// Device/Application/02_Devices/FB_RealCylinderGroup
FUNCTION_BLOCK FB_RealCylinderGroup
(* 模块说明：按料型选通的真实气缸组适配层（G2 侧挡用，300/450/600 三缸共用设备索引 10）。
   同一时刻只允许一个气缸下降，其余两个强制提升；回写与 FB_SimDevice 完全一致的接收/完成序号，
   使上层流程与互锁无需区分单缸、多缸或仿真。
   命令目标 lrTarget：0 = 三缸全部提升；300 / 450 / 600 = 对应料型气缸下降，其余两个提升。
   lrTarget 在 0..1 之间时按单缸旧语义映射：>0.5 视为「降到当前料型」，<=0.5 视为三缸全部提升。 *)
VAR_INPUT
	xUseReal : BOOL; (* TRUE 表示本编号由真实气缸组接管；FALSE 时三个阀全部失电且不响应任何命令。 *)
	xEnable : BOOL; (* 设备级使能，来自整机许可；FALSE 时阀失电并清序号。 *)
	xReset : BOOL; (* 故障复位上升沿；清锁存错误与序号。 *)
	xFaultHold : BOOL; (* 整机故障保持：TRUE 时三个阀立即失电，直到复位。 *)
	uiMaterialModel : UINT; (* 当前运行料型 300/450/600；旧语义 lrTarget>0.5 时降到本料型。 *)
	xSensorRetract1 : BOOL; (* 1 号缸（300）提升到位传感器原始电平，TRUE 表示该端有信号。 *)
	xSensorExtend1 : BOOL; (* 1 号缸（300）下降到位传感器原始电平。 *)
	xSensorRetract2 : BOOL; (* 2 号缸（450）提升到位传感器原始电平。 *)
	xSensorExtend2 : BOOL; (* 2 号缸（450）下降到位传感器原始电平。 *)
	xSensorRetract3 : BOOL; (* 3 号缸（600）提升到位传感器原始电平。 *)
	xSensorExtend3 : BOOL; (* 3 号缸（600）下降到位传感器原始电平。 *)
	xInvertSensors : BOOL; (* TRUE 表示六个传感器均为低电平有效，本层统一取反，不动上层。 *)
	xInvertValve : BOOL; (* TRUE 表示三个阀均为低电平使能；默认 FALSE，即高电平使能。 *)
	tSensorTimeout : TIME := T#3S; (* 六个传感器全部无信号达到该时间判为整组丢失，报 3004。 *)
	tTravelTimeout : TIME := T#10S; (* 命令发出后目标姿态未达成达到该时间判为动作超时，报 3005。 *)
	stConfig : ST_DeviceConfig; (* 行程范围，语义与仿真侧一致；组内气缸只使用 0/1 两端。 *)
	stCommand : ST_DeviceCommand; (* 上层统一设备命令，本层只响应 Position 的 0/300/450/600 目标。 *)
END_VAR
VAR_OUTPUT
	stStatus : ST_DeviceStatus; (* 与 FB_SimDevice 语义一致；目标缸下降到位 1.0，三缸全提 0.0，中间保持上次值。 *)
	aValve : ARRAY[1..3] OF BOOL; (* 三个阀的电气电平（已含 xInvertValve），直接接物理输出点；索引 1=300，2=450，3=600。 *)
	uiActiveBand : UINT; (* 当前实际下降的料型带号；0 表示三个缸都在提升位。 *)
END_VAR
VAR
	rtReset : R_TRIG; (* 复位上升沿。 *)
	tonNoSensor : TON; (* 六个传感器全部无信号的持续计时。 *)
	tonTravel : TON; (* 命令发出后等待到位的计时。 *)
	udiLastID : UDINT; (* 上次已接受的命令序号。 *)
	aRetract : ARRAY[1..3] OF BOOL; (* 取反处理后的三路提升信号。 *)
	aExtend : ARRAY[1..3] OF BOOL; (* 取反处理后的三路下降信号。 *)
	xAllRetract : BOOL; (* 三个缸都确认在提升位。 *)
	xPositionKnown : BOOL; (* 三缸姿态是否都已由传感器确立；未确立时 xReady 必须为 FALSE，防止上层把未知当成已提升。 *)
	xCmdValid : BOOL; (* 当前存在有效的保位命令，阀按此持续输出。 *)
	uiTargetBand : UINT; (* 有效命令期望下降的料型带号；0 表示三缸全部提升。 *)
	xTravelling : BOOL; (* 尚未确认到达命令要求的姿态。 *)
	i : INT; (* 本扫描数组遍历索引；含义及范围以当前 FOR 循环为准。 *)
END_VAR

rtReset(CLK := xReset);

(* ===== 1. 复位：只清错误与序号，姿态仍由传感器决定 ===== *)
IF xUseReal AND rtReset.Q THEN
	stStatus.xError := FALSE; stStatus.udiErrorID := 0;
	xCmdValid := FALSE; xTravelling := FALSE; udiLastID := 0; uiTargetBand := 0;
	stStatus.udiAcceptedID := 0; stStatus.udiCompletedID := 0;
	tonNoSensor(IN := FALSE);
	tonTravel(IN := FALSE);
END_IF

(* ===== 2. 传感器取反与逐缸姿态判定 ===== *)
aRetract[1] := xSensorRetract1 XOR xInvertSensors;
aExtend[1] := xSensorExtend1 XOR xInvertSensors;
aRetract[2] := xSensorRetract2 XOR xInvertSensors;
aExtend[2] := xSensorExtend2 XOR xInvertSensors;
aRetract[3] := xSensorRetract3 XOR xInvertSensors;
aExtend[3] := xSensorExtend3 XOR xInvertSensors;

(* 单缸两端同时有信号：传感器短路、磁环位置错或机械卡在中间，该缸姿态不可信，按 3003 暴露。
   逐缸判定而不是整组判定：只要有一个缸自相矛盾，整组位置就不可信。 *)
FOR i := 1 TO 3 DO
	IF aRetract[i] AND aExtend[i] THEN
		stStatus.xError := TRUE; stStatus.udiErrorID := 3003;
	END_IF
END_FOR

(* 三缸姿态是否都已确立：每个缸必须恰好一端有效，中间态或两端全无都算未确立。 *)
xAllRetract := aRetract[1] AND aRetract[2] AND aRetract[3];
xPositionKnown := TRUE;
FOR i := 1 TO 3 DO
	IF (NOT aRetract[i]) AND (NOT aExtend[i]) THEN xPositionKnown := FALSE; END_IF
END_FOR
IF stStatus.xError THEN xPositionKnown := FALSE; END_IF

(* 六个传感器全部无信号并持续 tSensorTimeout：判整组传感器丢失，报 3004。
   单缸丢失不在这里报，由 xPositionKnown 为 FALSE 阻断就绪，交给超时暴露，避免一缸调试刷整组报警。 *)
tonNoSensor(IN := xUseReal AND NOT aRetract[1] AND NOT aExtend[1]
	AND NOT aRetract[2] AND NOT aExtend[2]
	AND NOT aRetract[3] AND NOT aExtend[3], PT := tSensorTimeout);
IF tonNoSensor.Q AND NOT stStatus.xError THEN
	stStatus.xError := TRUE; stStatus.udiErrorID := 3004;
END_IF

(* ===== 3. 命令接收与保位判定 ===== *)
IF NOT xUseReal THEN
	(* 未接管：不驱动阀，也不发布就绪，避免被上层当成可用设备 *)
	xCmdValid := FALSE; xTravelling := FALSE; udiLastID := 0; uiTargetBand := 0;
	stStatus.xReady := FALSE; stStatus.xBusy := FALSE; stStatus.xActive := FALSE;
	stStatus.udiAcceptedID := 0; stStatus.udiCompletedID := 0;
ELSIF NOT xEnable OR stStatus.xError OR xFaultHold THEN
	(* 故障或整机故障保持时阀失电，不带错误继续动作 *)
	xCmdValid := FALSE; xTravelling := FALSE;
	stStatus.xReady := FALSE; stStatus.xBusy := FALSE; stStatus.xActive := FALSE;
ELSE
	stStatus.xReady := xEnable AND xPositionKnown;

	(* 新序号即新命令；姿态未确立时不接受，防止朝未知状态动作 *)
	IF (stCommand.udiID <> 0) AND (stCommand.udiID <> udiLastID)
		AND xEnable AND xPositionKnown AND NOT stStatus.xBusy THEN
		udiLastID := stCommand.udiID;
		stStatus.udiAcceptedID := udiLastID; stStatus.udiCompletedID := 0;
		CASE stCommand.eAction OF
		E_DeviceAction.Position:
			IF (stCommand.lrTarget > 0.5) AND (stCommand.lrTarget <= 1.0) THEN
				(* 单缸旧语义：1 = 降到当前料型；料型非法时报 2001，不猜一个缸去动作 *)
				IF (uiMaterialModel = 300) OR (uiMaterialModel = 450) OR (uiMaterialModel = 600) THEN
					uiTargetBand := uiMaterialModel;
				ELSE
					stStatus.xError := TRUE; stStatus.udiErrorID := 2001;
				END_IF
			ELSIF ABS(stCommand.lrTarget) < 0.01 THEN
				uiTargetBand := 0;
			ELSIF (ABS(stCommand.lrTarget - 300.0) < 0.01) THEN
				uiTargetBand := 300;
			ELSIF (ABS(stCommand.lrTarget - 450.0) < 0.01) THEN
				uiTargetBand := 450;
			ELSIF (ABS(stCommand.lrTarget - 600.0) < 0.01) THEN
				uiTargetBand := 600;
			ELSE
				(* 只支持 0 / 300 / 450 / 600，其它目标明确报错而不是静默不动 *)
				stStatus.xError := TRUE; stStatus.udiErrorID := 2001;
			END_IF
			IF NOT stStatus.xError THEN
				xCmdValid := TRUE;
				xTravelling := TRUE;
				stStatus.xBusy := TRUE;
			ELSE
				xCmdValid := FALSE;
			END_IF
		E_DeviceAction.Stop, E_DeviceAction.None:
			xCmdValid := FALSE; xTravelling := FALSE; uiTargetBand := 0;
			stStatus.udiAcceptedID := 0; stStatus.udiCompletedID := 0;
			udiLastID := 0;
		ELSE
			(* 气缸组没有连续运行、点动和回零，明确报错而不是静默不动 *)
			stStatus.xError := TRUE; stStatus.udiErrorID := 2001;
			xCmdValid := FALSE;
		END_CASE
	END_IF

	(* 命令被撤销或失能：立即取消保位，阀随之失电 *)
	IF (stCommand.eAction = E_DeviceAction.Stop) OR (stCommand.eAction = E_DeviceAction.None)
		OR NOT xEnable THEN
		xCmdValid := FALSE; xTravelling := FALSE;
		stStatus.xBusy := FALSE;
	END_IF

	(* 到位判定：目标缸下降到位，并且另外两个缸都在提升位，才算本次命令完成。
	   中间态（目标缸还没下去、或另一缸还没起来）都视为未完成，由超时兜底。 *)
	IF xCmdValid AND xPositionKnown THEN
		CASE uiTargetBand OF
		0:
			IF xAllRetract THEN
				IF xTravelling THEN stStatus.udiCompletedID := udiLastID; END_IF
				xTravelling := FALSE;
				stStatus.xBusy := FALSE;
			END_IF
		300:
			IF aExtend[1] AND aRetract[2] AND aRetract[3] THEN
				IF xTravelling THEN stStatus.udiCompletedID := udiLastID; END_IF
				xTravelling := FALSE;
				stStatus.xBusy := FALSE;
			END_IF
		450:
			IF aExtend[2] AND aRetract[1] AND aRetract[3] THEN
				IF xTravelling THEN stStatus.udiCompletedID := udiLastID; END_IF
				xTravelling := FALSE;
				stStatus.xBusy := FALSE;
			END_IF
		600:
			IF aExtend[3] AND aRetract[1] AND aRetract[2] THEN
				IF xTravelling THEN stStatus.udiCompletedID := udiLastID; END_IF
				xTravelling := FALSE;
				stStatus.xBusy := FALSE;
			END_IF
		END_CASE
	END_IF
END_IF

(* ===== 4. 位置反馈：只有确切在位才更新，中间态保持上次值 ===== *)
IF uiTargetBand = 0 THEN
	IF xAllRetract THEN stStatus.lrPosition := 0.0; END_IF
ELSIF uiTargetBand = 300 THEN
	IF aExtend[1] THEN stStatus.lrPosition := 1.0; END_IF
ELSIF uiTargetBand = 450 THEN
	IF aExtend[2] THEN stStatus.lrPosition := 1.0; END_IF
ELSIF uiTargetBand = 600 THEN
	IF aExtend[3] THEN stStatus.lrPosition := 1.0; END_IF
END_IF

(* 实际下降的料型：命令目标有效且该缸确实到位才报带号，避免阀已得电但没下去时谎报挡料就位 *)
uiActiveBand := 0;
IF (uiTargetBand = 300) AND aExtend[1] THEN uiActiveBand := 300; END_IF
IF (uiTargetBand = 450) AND aExtend[2] THEN uiActiveBand := 450; END_IF
IF (uiTargetBand = 600) AND aExtend[3] THEN uiActiveBand := 600; END_IF

(* ===== 5. 到位超时 ===== *)
tonTravel(IN := xUseReal AND xTravelling AND xCmdValid, PT := tTravelTimeout);
IF tonTravel.Q AND NOT stStatus.xError THEN
	stStatus.xError := TRUE; stStatus.udiErrorID := 3005;
	stStatus.xBusy := FALSE;
	xTravelling := FALSE;
END_IF

(* ===== 6. 阀输出：按保位命令持续输出，不是只在动作过程中输出；任何时刻最多一个缸下降 ===== *)
aValve[1] := FALSE; aValve[2] := FALSE; aValve[3] := FALSE;
IF xCmdValid AND xUseReal AND NOT stStatus.xError AND NOT xFaultHold THEN
	aValve[1] := (uiTargetBand = 300);
	aValve[2] := (uiTargetBand = 450);
	aValve[3] := (uiTargetBand = 600);
END_IF
IF xInvertValve THEN
	aValve[1] := NOT aValve[1]; aValve[2] := NOT aValve[2]; aValve[3] := NOT aValve[3];
END_IF

(* ===== 7. 收尾 ===== *)
stStatus.xReady := stStatus.xReady AND xUseReal AND NOT stStatus.xError;
stStatus.xActive := xCmdValid;
(* 气缸组没有回零动作，用「三缸姿态都已确立」代替，供整机统计已接管设备是否可信 *)
stStatus.xHomed := xUseReal AND xPositionKnown;

END_FUNCTION_BLOCK

// Device/Application/02_Devices/FB_RealSensor
FUNCTION_BLOCK FB_RealSensor
(* 模块说明：真实传感器（光电/接近开关）只读适配层。本块不驱动任何输出，只把原始电平
   去抖后发布成「到位」状态，使上层（自动送料判断、互锁、诊断）与仿真设备使用同一套接口。
   按料型/来料判断的是「有没有件」而不是「走到哪个位置」，所以姿态只有 0.0 / 1.0 两端：
   1.0 = 有料（光电被遮挡），0.0 = 无料。连续位置对传感器没有意义。 *)
VAR_INPUT
	xUseReal : BOOL; (* TRUE 表示本编号由真实传感器接管；FALSE 时不读物理点，也不发布就绪。 *)
	xEnable : BOOL; (* 设备级使能，来自整机许可；FALSE 时状态复位为无料且不发布就绪。 *)
	xReset : BOOL; (* 故障复位上升沿；清锁存错误。 *)
	xSensorRaw : BOOL; (* 传感器原始电平，TRUE 表示被遮挡（有料）。 *)
	xInvertSensor : BOOL; (* TRUE 表示接线为低电平有效（遮挡时读 FALSE），本层统一取反，不动上层。 *)
	tDebounce : TIME := T#20MS; (* 去抖时间：光电受粉尘、振动、反光影响会抖，短于该时间的跳变忽略。 *)
	tStuckTimeout : TIME := T#0MS; (* 常亮/常灭监视；0 表示不监视。料走完仍长时间有信号通常代表传感器卡死或反光。 *)
	stConfig : ST_DeviceConfig; (* 与其它设备一致的配置结构；传感器只用 lrInitialPosition 作初值，不使用行程字段。 *)
	stCommand : ST_DeviceCommand; (* 上层统一设备命令；传感器只响应被读请求，Position 目标被忽略。 *)
END_VAR
VAR_OUTPUT
	stStatus : ST_DeviceStatus; (* 与仿真侧语义一致；lrPosition 取 1.0 有料、0.0 无料。 *)
	xDetected : BOOL; (* 去抖后的最终信号，TRUE=有料。流程与互锁直接取用这个而不是原始点。 *)
	xRaw : BOOL; (* 取反处理后的原始电平（未去抖），供在线排查接线极性与抖动。 *)
END_VAR
VAR
	rtReset : R_TRIG; (* 复位上升沿。 *)
	tonDebounce : TON; (* 由 FALSE 变 TRUE 的去抖计时，到时才认「有料」。 *)
	tonClear : TON; (* 由 TRUE 变 FALSE 的去抖计时，到时才认「无料」。 *)
	tonStuck : TON; (* 长时间保持同一状态计时，用于常亮/常灭监视。 *)
	xStuckWindowClear : BOOL; (* 本扫描检测到电平跳变：清掉常亮/常灭计时窗口，重新开始计时。 *)
	xStable : BOOL; (* 去抖后的稳定值。 *)
	xLastRaw : BOOL; (* 上扫描取反后的原始电平，用于判断是否发生跳变并重置去抖计时。 *)
	xBooted : BOOL; (* 首次扫描标志，上电时直接用当前电平作初值，不等待去抖。 *)
END_VAR

rtReset(CLK := xReset);

(* ===== 1. 复位：只清错误，状态仍由传感器决定 ===== *)
IF xUseReal AND rtReset.Q THEN
	stStatus.xError := FALSE; stStatus.udiErrorID := 0;
	tonStuck(IN := FALSE);
END_IF

(* ===== 2. 极性处理：接线反了只改 xInvertSensor 一个参数，上层不受影响 ===== *)
xRaw := xSensorRaw XOR xInvertSensor;

(* ===== 3. 去抖：跳变后必须稳定 tDebounce 才改 xStable ===== *)
(* 用两个单稳计时而不是一个沿检测，是为了让"抖动期间保持上次稳定值"这件事显式可见：
   信号连续抖动时两个计时都不会到时，xStable 保持在最后一个稳定值上。 *)
xStuckWindowClear := (NOT xBooted) OR (xRaw <> xLastRaw);
IF xStuckWindowClear THEN
	tonDebounce(IN := FALSE);
	tonClear(IN := FALSE);
	IF NOT xBooted THEN
		(* 上电直接用当前电平作初值，避免开机 20ms 内把有料当无料 *)
		xStable := xRaw;
		xBooted := TRUE;
	END_IF
	xLastRaw := xRaw;
END_IF

IF xUseReal THEN
	IF xRaw THEN
		tonDebounce(IN := TRUE, PT := tDebounce);
		tonClear(IN := FALSE);
		IF tonDebounce.Q THEN xStable := TRUE; END_IF
	ELSE
		tonClear(IN := TRUE, PT := tDebounce);
		tonDebounce(IN := FALSE);
		IF tonClear.Q THEN xStable := FALSE; END_IF
	END_IF
END_IF

xDetected := xStable;

(* ===== 4. 常亮/常灭监视：料已走完却一直有信号，或本该有料却一直没有，都报出来 =====
   只监视"信号纹丝不动"这个可观测事实，不猜业务含义；阈值由 tStuckTimeout 给，0 表示关闭。 *)
tonStuck(IN := xUseReal AND (tStuckTimeout > T#0MS) AND NOT xStuckWindowClear, PT := tStuckTimeout);
IF tonStuck.Q AND NOT stStatus.xError THEN
	stStatus.xError := TRUE;
	(* 3006：持续有信号（常亮/反光/卡死）；3007：持续无信号（断线/被挡/未接通） *)
	IF xDetected THEN stStatus.udiErrorID := 3006;
	ELSE stStatus.udiErrorID := 3007; END_IF
END_IF

(* ===== 5. 状态发布：传感器没有动作请求，只要接管且使能就算就绪 ===== *)
stStatus.lrPosition := SEL(xDetected, 0.0, 1.0);
stStatus.xReady := xUseReal AND xEnable AND NOT stStatus.xError;
stStatus.xActive := xUseReal AND xDetected;
stStatus.xBusy := FALSE;
(* 传感器没有回零概念，用"已接管且状态可信"代替 *)
stStatus.xHomed := xUseReal AND xBooted;
stStatus.xRealActive := xUseReal;

END_FUNCTION_BLOCK

// Device/Application/04_Machine/FB_ManualControl
(* 模块说明：将手动按钮转为统一设备请求。点动松开即取消；定位与回零请求保持到本次完成；D6 不调度。 *)
FUNCTION_BLOCK FB_ManualControl
VAR_INPUT
	xEnable : BOOL; (* 手动模式且按钮释放联锁已满足时允许；未使能也同步按钮快照。 *)
	stReal : ST_RealDeviceSettings; (* 真实设备接管设置；真实编号的手动速度收紧到验证速度。 *)
	aManual : ARRAY[1..17] OF ST_ManualCommand; (* 各设备手动请求，索引 1..17；进入手动后先释放所有按钮再允许动作。 *)
END_VAR
VAR_IN_OUT
	aCommand : ARRAY[1..17] OF ST_DeviceCommand; (* 统一设备请求数组 1..17；子流程写请求，设备管理器执行。 *)
	aStatus : ARRAY[1..17] OF ST_DeviceStatus; (* 各设备的反馈数组 1..17，供判断忙、完成序号、故障和位置。 *)
	udiCounter : UDINT; (* 全机共享的动作序号计数器，通过引用传递；由 F_NextID 分配，0 不使用。 *)
END_VAR
VAR_OUTPUT
	uiRejectDevice : UINT; (* 本扫描最后一个手动拒绝设备索引；0 无，常见原因是冲突按钮或不支持该动作。 *)
END_VAR
VAR
	aPrev : ARRAY[1..17] OF ST_ManualCommand; (* 上扫描手动按钮快照；即使禁用仍更新，防止按住按钮切模式后被误作新上升沿。 *)
	aPending : ARRAY[1..17] OF ST_DeviceCommand; (* 手动定位或回零的锁存请求，直到本次命令完成；点动或运行优先时清除。 *)
	aRunID : ARRAY[1..17] OF UDINT; (* 各设备按住运行/点动时保持的序号，按钮释放后归零。 *)
	i : INT; (* 本扫描数组遍历索引；含义及范围以当前 FOR 循环为准。 *)
	lrVelocity : LREAL; (* 本扫描限幅后的手动速度，取绝对值限幅 0.1..100；反向点动时变为负值。 *)
	lrVelocityMax : LREAL; (* 本扫描速度上限；真实设备收紧到验证速度，防止全速冲出。 *)
	uiPressed : UINT; (* 本扫描该设备同时按下的手动按钮个数；大于 1 视为冲突并拒绝。 *)
END_VAR

(* 每扫描重新判断按钮冲突；无合法请求的设备由整机统一撤销动作。 *)
uiRejectDevice:=0;
FOR i:=1 TO 17 DO
    IF NOT xEnable THEN
        aPending[i].eAction:=E_DeviceAction.None;
        aRunID[i]:=0;
    ELSIF i<>6 THEN
        (* 先撤销本设备请求，只有命中合法按钮时才在下面重新写入。否则松开点动后，
           上一扫描的 Jog 会一直残留在共享请求数组里，真实轴靠 None/Stop 停止的逻辑永远等不到。 *)
        aCommand[i]:=F_Command(E_DeviceAction.None,0,0.0,0.0);
        (* 真实设备的手动速度上限由 lrManualVelocityMax 决定（默认 200）；实际速度取 aManual[i].lrVelocity 与之较小者。 *)
        lrVelocityMax:=100.0;
        IF stReal.axRealDevice[i] THEN
            (* 新字段在未重新初始化的旧下载里可能为 0；兜底 100，避免手动速度变 0 表现为不动作 *)
            lrVelocityMax:=100.0;
            IF stReal.lrManualVelocityMax>0.1 THEN lrVelocityMax:=LIMIT(0.1,stReal.lrManualVelocityMax,200.0); END_IF
        END_IF
        IF i=8 THEN
            (* D8 平台旋转轴（主轴）手动默认 3、限速 5；请求值超过上限时按默认 3 走，不要直接跳到 5。 *)
            lrVelocityMax:=5.0;
            lrVelocity:=3.0;
            IF ABS(aManual[i].lrVelocity)<=lrVelocityMax THEN
                lrVelocity:=LIMIT(0.1,ABS(aManual[i].lrVelocity),lrVelocityMax);
            END_IF
        ELSE
            lrVelocity:=LIMIT(0.1,ABS(aManual[i].lrVelocity),lrVelocityMax);
        END_IF
        (* 任意两个手动按钮同时按下都算冲突：正反点动、点动与定位/运行/回零、定位与运行/回零、运行与回零。 *)
        uiPressed:=0;
        IF aManual[i].xJogPositive THEN uiPressed:=uiPressed+1; END_IF
        IF aManual[i].xJogNegative THEN uiPressed:=uiPressed+1; END_IF
        IF aManual[i].xMove THEN uiPressed:=uiPressed+1; END_IF
        IF aManual[i].xRun THEN uiPressed:=uiPressed+1; END_IF
        IF aManual[i].xHome THEN uiPressed:=uiPressed+1; END_IF
        IF uiPressed>1 THEN
            uiRejectDevice:=INT_TO_UINT(i); aPending[i].eAction:=E_DeviceAction.None;
        (* 点动电平控制，只支持 D2/D4/D5/D7/D8；速度符号决定方向，松开后不保持点动。 *)
        ELSIF aManual[i].xJogPositive OR aManual[i].xJogNegative THEN
            aPending[i].eAction:=E_DeviceAction.None;
            IF aRunID[i]=0 THEN aRunID[i]:=F_NextID(udiCounter); END_IF
            IF aManual[i].xJogNegative THEN lrVelocity:=-lrVelocity; END_IF
            IF (i=2) OR (i=4) OR (i=5) OR (i=7) OR (i=8) THEN
                aCommand[i]:=F_Command(E_DeviceAction.Jog,aRunID[i],0.0,lrVelocity);
            ELSE uiRejectDevice:=INT_TO_UINT(i);
            END_IF
        (* 连续运行电平控制，仅允许皮带、盘刀、喷油和吹气；盘刀接真实轴后走 FB_RealAxis 的 Run 相位。 *)
        ELSIF aManual[i].xRun THEN
            aPending[i].eAction:=E_DeviceAction.None;
            IF (i=1) OR (i=3) OR (i=13) OR (i=14) THEN
                IF aRunID[i]=0 THEN aRunID[i]:=F_NextID(udiCounter); END_IF
                aCommand[i]:=F_Command(E_DeviceAction.Run,aRunID[i],0.0,lrVelocity);
            ELSE uiRejectDevice:=INT_TO_UINT(i);
            END_IF
        (* 回零：上升沿锁存一次请求，之后每扫描重发直到完成；真实轴 D2/D8，D4 为仿真但保留入口。
           D3 盘刀是连续旋转主轴，只做 Run 不做回零，因此不在本白名单内。
           这里不能像点动那样在分支开头清 aPending —— 回零是保持型动作，清了就只剩一个扫描周期，
           设备刚接收就会被下一扫描的 None 撤销，表现为「下发了但不动」。 *)
        ELSIF aManual[i].xHome THEN
            aRunID[i]:=0;
            IF (i=2) OR (i=4) OR (i=8) THEN
                IF NOT aPrev[i].xHome THEN
                    aPending[i]:=F_Command(E_DeviceAction.Home,F_NextID(udiCounter),0.0,0.0);
                END_IF
                IF aPending[i].eAction<>E_DeviceAction.None THEN
                    aCommand[i]:=aPending[i];
                    IF F_Done(aStatus[i],aPending[i].udiID) THEN aPending[i].eAction:=E_DeviceAction.None; END_IF
                END_IF
            ELSE
                (* 不支持的编号：清掉可能从定位继承来的请求，避免继续执行上一个动作。 *)
                uiRejectDevice:=INT_TO_UINT(i);
                aPending[i].eAction:=E_DeviceAction.None;
            END_IF
        ELSE
            aRunID[i]:=0;
            (* 定位仅在按钮上升沿锁存目标和序号，然后持续等待本次完成。 *)
            IF aManual[i].xMove AND NOT aPrev[i].xMove THEN
                IF (i<>1) AND (i<>3) AND (i<>13) AND (i<>14) THEN
                    aPending[i]:=F_Command(E_DeviceAction.Position,F_NextID(udiCounter),aManual[i].lrTarget,lrVelocity);
                ELSE uiRejectDevice:=INT_TO_UINT(i);
                END_IF
            END_IF
            IF aPending[i].eAction<>E_DeviceAction.None THEN
                aCommand[i]:=aPending[i];
                IF F_Done(aStatus[i],aPending[i].udiID) THEN aPending[i].eAction:=E_DeviceAction.None; END_IF
            END_IF
        END_IF
    END_IF
    (* 禁用时仍同步按钮快照，避免按住定位按钮切入手动后产生虚假的新上升沿。 *)
    aPrev[i]:=aManual[i];
END_FOR

END_FUNCTION_BLOCK

// Device/Application/02_Devices/F_Command
(* 模块说明：组装设备命令，不执行运动。由设备管理器和对应设备功能块实际处理。 *)
FUNCTION F_Command : ST_DeviceCommand
VAR_INPUT
    eAction : E_DeviceAction; (* 动作类型：无请求、定位、连续运行、点动或停止，见 E_DeviceAction。 *)
    udiID : UDINT; (* 本次命令序号，0 无效；发起新定位时换新序号。 *)
    lrTarget : LREAL; (* 目标工程位置；气缸使用约定的 0/1 端点，连续运行和点动不使用该位置。 *)
    lrVelocity : LREAL; (* 请求速度，单位随设备工程单位定义；尚未完成实机标定。 *)
END_VAR

(* 只复制字段形成结构体，不等待动作、不直接访问物理设备。 *)
F_Command.eAction := eAction;
F_Command.udiID := udiID;
F_Command.lrTarget := lrTarget;
F_Command.lrVelocity := lrVelocity;

END_FUNCTION

// Device/Application/02_Devices/F_NextID
(* 模块说明：生成本次动作的非零序号。计数到最大值后回到 1，用于排除上一步残留的完成反馈。 *)
FUNCTION F_NextID : UDINT
VAR_IN_OUT
    udiCounter : UDINT; (* 全机共享的动作序号计数器，通过引用传递；由 F_NextID 分配，0 不使用。 *)
END_VAR

(* 最大值之后回到 1，跳过无效序号 0；同一机台所有流程共享该计数器。 *)
IF udiCounter = 16#FFFFFFFF THEN udiCounter := 1;
ELSE udiCounter := udiCounter + 1;
END_IF
F_NextID := udiCounter;

END_FUNCTION

// Device/Application/02_Devices/F_Done
(* 模块说明：只有设备完成序号等于本次命令序号、无忙且无故障，才返回动作完成。 *)
FUNCTION F_Done : BOOL
VAR_INPUT
    stStatus : ST_DeviceStatus; (* 本模块对外发布的状态；字段含义见其数据类型。 *)
    udiID : UDINT; (* 本次命令序号，0 无效；发起新定位时换新序号。 *)
END_VAR

(* 完成必须匹配本次请求；历史 Done 或仅 Busy=FALSE 都不足以作为本步完成条件。 *)
F_Done := (udiID <> 0) AND (stStatus.udiCompletedID = udiID)
    AND NOT stStatus.xBusy AND NOT stStatus.xError;

END_FUNCTION

// Device/Application/04_Machine/FB_AutoCycle
(* 模块说明：自动主状态机。只组织工序并提出请求，设备执行由整机统一调用；送料等料允许长期等待。 *)
FUNCTION_BLOCK FB_AutoCycle
VAR_INPUT
    xRun : BOOL; (* 自动工序运行许可，整机 Automatic 时保持 TRUE；撤销立即复位主流程。 *)
    xContinuous : BOOL; (* TRUE 连续循环；FALSE 在当前完整循环结束后回到就绪。 *)
    xMaterialAtLength : BOOL; (* 定长光电到位状态；自动送料须先离开再到位，并满足 D5 下降。 *)
    stRecipe : ST_Recipe; (* 待校验配方或上层传入的运行配方，字段含义见 ST_Recipe。 *)
END_VAR
VAR_IN_OUT
    aCommand : ARRAY[1..17] OF ST_DeviceCommand; (* 统一设备请求数组 1..17；子流程写请求，设备管理器执行。 *)
    aStatus : ARRAY[1..17] OF ST_DeviceStatus; (* 各设备的反馈数组 1..17，供判断忙、完成序号、故障和位置。 *)
    udiCounter : UDINT; (* 全机共享的动作序号计数器，通过引用传递；由 F_NextID 分配，0 不使用。 *)
END_VAR
VAR_OUTPUT
    eStep : E_AutoStep; (* 自动主工序当前状态，见 E_AutoStep。 *)
    xDone : BOOL; (* 整循环完成的单扫描脉冲；机械手等三路收尾全部结束后才产生。 *)
    xError : BOOL; (* 本设备或本子流程发生故障；具体原因见对应错误码。 *)
    udiErrorID : UDINT; (* 非法主步骤为 4800；主步超时为 4800+步号；步骤守护失败为 4800+步号+1，见下方守护表；支线错误则向上传递。 *)
    uiClearLengthStep : UINT; (* 避让支线 P 的当前步骤：10 升起 D5，20 移开 D4，1000 完成。 *)
    uiClearTransferStep : UINT; (* 避让支线 Q 当前步骤：10 降 G4，20 松 G3，30 降 G2，1000 完成。 *)
    uiPostStep : UINT; (* 收尾总步骤：10 抬刀，20 抬压，30 等待三路完成，1000 结束。 *)
    uiReturnKnifeStep : UINT; (* 收尾支线 A：10 喷油，20 D2 回刀，1000 完成。 *)
    uiUnloadStep : UINT; (* 机械手移料支线 B 步骤，10..110 每步加 10，1000 完成；详见 FB_Unload。 *)
    uiResetLengthStep : UINT; (* 收尾支线 C：10 D4 定位，20 D5 下降，30 确认下降，1000 完成。 *)
END_VAR
VAR
    ePrevStep : E_AutoStep := E_AutoStep.Fault; (* 上扫描主工序状态，用于产生步骤入口标志。 *)
    udiToken : UDINT; (* 本步骤专用动作序号；同一步中的设备共用该号，以排除旧完成信号。 *)
    udiSpindleToken : UDINT; (* 盘刀运行命令序号，切割过程中保持该号，避免重复重启盘刀命令。 *)
    udiPressToken : UDINT; (* G1 下压保位序号；PressDown 入口分配，后续步骤持续用该号重发，保证单电控阀不断电。 *)
    udiKnifeToken : UDINT; (* G9 下刀保位序号；KnifeDown 入口分配，同上。 *)
    xEntry : BOOL; (* 本扫描为新步骤入口；用于分配新序号并复位步骤超时计时。 *)
    xSawSensorClear : BOOL; (* 本轮送料已观察到光电离开；须先有该标志再接受新到位，防止残留信号触发。 *)
    tonStep : TON; (* 步骤超时定时器；进入新步骤时复位，超时错误码由模块及当前步号组成。 *)
    tStepLimit : TIME; (* 本扫描用的步骤超时值：切割步取 tCutTimeout，其余取 tStepTimeout。 *)
    xGuardOK : BOOL; (* 步骤守护判据：当前步依赖的前提是否仍满足，FALSE 时立即报错退出，不等步超时。 *)
    fbClear : FB_ClearanceUnit; (* 切割前两路并行避让流程。 *)
    fbPost : FB_PostCut; (* 切割后抬刀、抬压及三路收尾流程。 *)
END_VAR

(* 完成标志每扫描先清零；本流程在许可撤销后复位，不保留中断点续跑。 *)
xDone := FALSE;
IF NOT xRun THEN eStep:=E_AutoStep.Idle; xError:=FALSE; udiErrorID:=0; xSawSensorClear:=FALSE; END_IF
(* 进入新步骤才换新动作序号，同一步持续保持请求，防止反复启动。 *)
xEntry := eStep <> ePrevStep;
IF xEntry THEN udiToken := F_NextID(udiCounter); END_IF
ePrevStep := eStep;
(* 送料等料不计步骤超时；其余执行步按运行配方监控。
   切割步单独用 tCutTimeout：走刀行程长，和其它单动作步共用一个 30 秒很容易误超时。 *)
tStepLimit := stRecipe.tStepTimeout;
IF eStep = E_AutoStep.Cutting THEN tStepLimit := stRecipe.tCutTimeout; END_IF
tonStep(IN:=xRun AND NOT xEntry AND (eStep<>E_AutoStep.Idle)
    AND (eStep<>E_AutoStep.FeedWait) AND (eStep<>E_AutoStep.Complete)
    AND (eStep<>E_AutoStep.Fault),PT:=tStepLimit);
IF xRun AND NOT xError THEN
CASE eStep OF
(* 待机转入送料；没有直接跳到切割。 *)
E_AutoStep.Idle: eStep:=E_AutoStep.FeedWait;
(* D1 送料并正常等料；光电须先离开再到位，且 D5 必须在下降端。 *)
E_AutoStep.FeedWait:
    IF xEntry THEN xSawSensorClear:=FALSE; END_IF
    IF NOT xMaterialAtLength THEN xSawSensorClear:=TRUE; END_IF
    aCommand[1]:=F_Command(E_DeviceAction.Run,udiToken,0.0,stRecipe.lrBeltVelocity);
    IF xSawSensorClear AND xMaterialAtLength AND F_At(aStatus[5],1.0) THEN eStep:=E_AutoStep.StopFeed; END_IF
(* 本步不再给 D1 运行请求，整机周期清空请求后等待皮带非运行、非忙。 *)
E_AutoStep.StopFeed:
    IF NOT aStatus[1].xActive AND NOT aStatus[1].xBusy THEN eStep:=E_AutoStep.Push; END_IF
(* G3 侧推到位；只认本次 udiToken 对应的完成。 *)
E_AutoStep.Push:
    aCommand[11]:=F_Command(E_DeviceAction.Position,udiToken,1.0,stRecipe.lrPositionVelocity);
    IF F_Done(aStatus[11],udiToken) THEN eStep:=E_AutoStep.Clearance; END_IF
(* 并行调用定长避让 P 和输送机构避让 Q，两路都完成后旋转平台。 *)
E_AutoStep.Clearance:
    IF fbClear.xDone THEN eStep:=E_AutoStep.Rotate; END_IF
(* D8 旋转到 lrRotateAngle，必须在 G1 下压之前完成。 *)
E_AutoStep.Rotate:
    aCommand[8]:=F_Command(E_DeviceAction.Position,udiToken,stRecipe.lrRotateAngle,stRecipe.lrPositionVelocity);
    IF F_Done(aStatus[8],udiToken) THEN eStep:=E_AutoStep.PressDown; END_IF
(* G1 下压到位。 *)
E_AutoStep.PressDown:
    IF xEntry THEN udiPressToken:=udiToken; END_IF
    aCommand[9]:=F_Command(E_DeviceAction.Position,udiPressToken,1.0,stRecipe.lrPositionVelocity);
    IF F_Done(aStatus[9],udiPressToken) THEN eStep:=E_AutoStep.SpindleOn; END_IF
(* D3 盘刀先转起来，转稳了再下刀；此时刀还没下来，G1 保持压紧。 *)
E_AutoStep.SpindleOn:
    udiSpindleToken:=udiToken;
    aCommand[9]:=F_Command(E_DeviceAction.Position,udiPressToken,1.0,stRecipe.lrPositionVelocity);
    aCommand[3]:=F_Command(E_DeviceAction.Run,udiSpindleToken,0.0,stRecipe.lrSpindleVelocity);
    IF F_Done(aStatus[3],udiSpindleToken) AND aStatus[3].xActive THEN eStep:=E_AutoStep.KnifeDown; END_IF
(* G9 盘刀下降到位；下降全程 D3 保持运行。 *)
E_AutoStep.KnifeDown:
    IF xEntry THEN udiKnifeToken:=udiToken; END_IF
    aCommand[9]:=F_Command(E_DeviceAction.Position,udiPressToken,1.0,stRecipe.lrPositionVelocity);
    aCommand[3]:=F_Command(E_DeviceAction.Run,udiSpindleToken,0.0,stRecipe.lrSpindleVelocity);
    aCommand[17]:=F_Command(E_DeviceAction.Position,udiKnifeToken,1.0,stRecipe.lrPositionVelocity);
    IF F_Done(aStatus[17],udiKnifeToken) THEN eStep:=E_AutoStep.Cutting; END_IF
(* 保持 D3 运行，G6 吹气，D2 走到回刀起点加切割长度；以 D2 到位作为切割完成。 *)
E_AutoStep.Cutting:
    aCommand[9]:=F_Command(E_DeviceAction.Position,udiPressToken,1.0,stRecipe.lrPositionVelocity);
    aCommand[17]:=F_Command(E_DeviceAction.Position,udiKnifeToken,1.0,stRecipe.lrPositionVelocity);
    aCommand[3]:=F_Command(E_DeviceAction.Run,udiSpindleToken,0.0,stRecipe.lrSpindleVelocity);
    aCommand[14]:=F_Command(E_DeviceAction.Run,udiToken,0.0,0.0);
    aCommand[2]:=F_Command(E_DeviceAction.Position,udiToken,stRecipe.lrCutHome+stRecipe.lrCutLength,stRecipe.lrCutVelocity);
    IF F_Done(aStatus[2],udiToken) THEN eStep:=E_AutoStep.StopCut; END_IF
(* 撤销 D3/G6 运行请求，等待盘刀停止且吹气关闭后收尾。 *)
E_AutoStep.StopCut:
    aCommand[9]:=F_Command(E_DeviceAction.Position,udiPressToken,1.0,stRecipe.lrPositionVelocity);
    aCommand[17]:=F_Command(E_DeviceAction.Position,udiKnifeToken,1.0,stRecipe.lrPositionVelocity);
    IF NOT aStatus[3].xActive AND NOT aStatus[3].xBusy AND NOT aStatus[14].xActive THEN eStep:=E_AutoStep.PostCut; END_IF
(* 先抬刀再抬压，随后三支线同步执行；全部结束才完成本轮。 *)
E_AutoStep.PostCut:
    IF fbPost.xDone THEN eStep:=E_AutoStep.Complete; END_IF
(* 只在进入本步时输出一次完成脉冲；连续模式返回送料，单循环由整机回到 Ready。 *)
E_AutoStep.Complete:
    xDone:=xEntry;
    IF xContinuous THEN eStep:=E_AutoStep.FeedWait; END_IF
(* 保留流程错误状态；整机退出自动后才复位此流程。 *)
E_AutoStep.Fault: xError:=TRUE;
ELSE xError:=TRUE; udiErrorID:=4800;
END_CASE
(* ===== 步骤守护表 =====
   只判前提，不判目标：目标是本步自己要去达成的东西，由各步的 F_Done 判完成；
   这里判的是这一步所依赖的前提还在不在。前提在进入该步时就已成立，
   之后必须一直保持，一旦丢失立即报错退出，不再干等 tonStep 超时才发现。
   每个步骤都要在下面有明确交代，无守护也要写出来，避免以后分不清
   是真的不需要还是漏掉了。新增步骤时先到这里补一行。
   错误码约定：4800 + 步号 + 1，例 SpindleOn=4881、Cutting=4891。
   这里不主动发 Stop：报错后本流程转 Fault，下一扫描不再提出任何请求，
   设备管理器收到 None 即停止，轴走 MC_Stop，气缸阀失电。 *)
xGuardOK := TRUE;
CASE eStep OF
(* 无守护：要么在等外部条件，要么本步本身就在建立条件。 *)
E_AutoStep.Idle, E_AutoStep.FeedWait, E_AutoStep.StopFeed,
E_AutoStep.Push, E_AutoStep.Clearance, E_AutoStep.Rotate,
E_AutoStep.PressDown, E_AutoStep.StopCut,
E_AutoStep.PostCut, E_AutoStep.Complete, E_AutoStep.Fault:
    xGuardOK := TRUE;

(* 起盘刀前：只要已压紧；此时刀还没下来，不判下刀。 *)
E_AutoStep.SpindleOn:
    xGuardOK := F_At(aStatus[9],1.0);

(* 下刀期间：压紧且盘刀必须已经在转，不能拿一把没转的刀往下扎。 *)
E_AutoStep.KnifeDown:
    xGuardOK := F_At(aStatus[9],1.0) AND aStatus[3].xActive;

(* 切割全程：压紧、下刀、盘刀运行三者都必须保持。 *)
E_AutoStep.Cutting:
    xGuardOK := F_At(aStatus[9],1.0) AND F_At(aStatus[17],1.0) AND aStatus[3].xActive;
END_CASE
IF NOT xGuardOK THEN
    xError := TRUE;
    udiErrorID := 4800 + TO_UDINT(eStep) + 1;
END_IF
IF tonStep.Q THEN xError:=TRUE; udiErrorID:=4800+TO_UDINT(eStep); END_IF
END_IF
(* 子功能块必须每扫描调用，包括失能时复位；上方状态判断看到的是此前反馈。 *)
fbClear(xExecute:=xRun AND (eStep=E_AutoStep.Clearance),stRecipe:=stRecipe,aCommand:=aCommand,aStatus:=aStatus,udiCounter:=udiCounter);
fbPost(xExecute:=xRun AND (eStep=E_AutoStep.PostCut),stRecipe:=stRecipe,aCommand:=aCommand,aStatus:=aStatus,udiCounter:=udiCounter);
(* 任一支线错误向主流程上报；所有设备请求还须经过整机统一互锁。 *)
IF fbClear.xError OR fbPost.xError THEN xError:=TRUE; udiErrorID:=MAX(fbClear.udiErrorID,fbPost.udiErrorID); END_IF
IF xError THEN eStep:=E_AutoStep.Fault; END_IF
uiClearLengthStep:=fbClear.uiLengthStep; uiClearTransferStep:=fbClear.uiTransferStep;
uiPostStep:=fbPost.uiStep; uiReturnKnifeStep:=fbPost.uiKnifeStep;
uiUnloadStep:=fbPost.uiUnloadStep; uiResetLengthStep:=fbPost.uiLengthStep;

END_FUNCTION_BLOCK

// Device/Application/03_Units/FB_Unload
(* 模块说明：收尾支线 B：机械手移料。后退、下降、最终回位是三个独立动作，全部完成后才允许下一轮送料。 *)
FUNCTION_BLOCK FB_Unload
VAR_INPUT
    xExecute : BOOL; (* 子流程执行许可；须保持到完成，清 FALSE 复位该流程步骤和错误。 *)
    stRecipe : ST_Recipe; (* 待校验配方或上层传入的运行配方，字段含义见 ST_Recipe。 *)
END_VAR
VAR_IN_OUT
    aCommand : ARRAY[1..17] OF ST_DeviceCommand; (* 统一设备请求数组 1..17；子流程写请求，设备管理器执行。 *)
    aStatus : ARRAY[1..17] OF ST_DeviceStatus; (* 各设备的反馈数组 1..17，供判断忙、完成序号、故障和位置。 *)
    udiCounter : UDINT; (* 全机共享的动作序号计数器，通过引用传递；由 F_NextID 分配，0 不使用。 *)
END_VAR
VAR_OUTPUT
    xDone : BOOL; (* 本子流程完成标志；执行许可撤销后复位。 *)
    xError : BOOL; (* 本设备或本子流程发生故障；具体原因见对应错误码。 *)
    udiErrorID : UDINT; (* 非法步骤码 4400；动作超时码=4400+uiStep，可据此定位本支线等待点。 *)
    uiStep : UINT; (* 当前子步骤：0 待机，10/20/... 执行动作，1000 完成；切勿在线强制跳步。 *)
END_VAR
VAR
    uiPrevStep : UINT := 65535; (* 上扫描步骤，用于判断本扫描是否刚进入新步骤。 *)
    udiToken : UDINT; (* 本步骤专用动作序号；同一步中的设备共用该号，以排除旧完成信号。 *)
    xEntry : BOOL; (* 本扫描为新步骤入口；用于分配新序号并复位步骤超时计时。 *)
    tonStep : TON; (* 步骤超时定时器；进入新步骤时复位，超时错误码由模块及当前步号组成。 *)
    tonSpray : TON; (* 通用子流程模板的喷油定时器，只有 FB_ReturnKnife 用其完成条件。 *)
END_VAR

(* 执行许可撤销即复位；步骤入口换新序号，每步等待本次动作完成，超时码=模块基码+步号。 *)
IF NOT xExecute THEN uiStep := 0; xError := FALSE; udiErrorID := 0; END_IF;
xEntry := uiStep <> uiPrevStep;
IF xEntry THEN udiToken := F_NextID(udiCounter); END_IF;
uiPrevStep := uiStep;
tonStep(IN := xExecute AND (uiStep > 0) AND (uiStep < 1000) AND NOT xEntry, PT := stRecipe.tStepTimeout);
tonSpray(IN := xExecute AND (uiStep = 10) AND aStatus[13].xActive, PT := stRecipe.tSpray);
IF xExecute AND NOT xError THEN
CASE uiStep OF
0: (* 待机；许可有效时进入首个动作。 *) uiStep := 10;
10: (* B010 侧挡 G2 提升。 *)
aCommand[10] := F_Command(E_DeviceAction.Position, udiToken, 0.0, stRecipe.lrPositionVelocity);
IF F_Done(aStatus[10], udiToken) THEN uiStep := 20; END_IF;
20: (* B020 流利条 G4 提升。 *)
aCommand[12] := F_Command(E_DeviceAction.Position, udiToken, 1.0, stRecipe.lrPositionVelocity);
IF F_Done(aStatus[12], udiToken) THEN uiStep := 30; END_IF;
30: (* B030 机械手 G7 提升。 *)
aCommand[15] := F_Command(E_DeviceAction.Position, udiToken, 1.0, stRecipe.lrPositionVelocity);
IF F_Done(aStatus[15], udiToken) THEN uiStep := 40; END_IF;
40: (* B040 夹爪 G8 打开，准备前进取料。 *)
aCommand[16] := F_Command(E_DeviceAction.Position, udiToken, 0.0, stRecipe.lrPositionVelocity);
IF F_Done(aStatus[16], udiToken) THEN uiStep := 50; END_IF;
50: (* B050 机械手 D7 前进到取料位置 lrGripperFront。 *)
aCommand[7] := F_Command(E_DeviceAction.Position, udiToken, stRecipe.lrGripperFront, stRecipe.lrPositionVelocity);
IF F_Done(aStatus[7], udiToken) THEN uiStep := 60; END_IF;
60: (* B060 夹爪 G8 夹紧，确认后才拉料。 *)
aCommand[16] := F_Command(E_DeviceAction.Position, udiToken, 1.0, stRecipe.lrPositionVelocity);
IF F_Done(aStatus[16], udiToken) THEN uiStep := 70; END_IF;
70: (* B070 机械手 D7 拉料到 lrGripperPull。 *)
aCommand[7] := F_Command(E_DeviceAction.Position, udiToken, stRecipe.lrGripperPull, stRecipe.lrPositionVelocity);
IF F_Done(aStatus[7], udiToken) THEN uiStep := 80; END_IF;
80: (* B080 夹爪 G8 打开，释放移走的料。 *)
aCommand[16] := F_Command(E_DeviceAction.Position, udiToken, 0.0, stRecipe.lrPositionVelocity);
IF F_Done(aStatus[16], udiToken) THEN uiStep := 90; END_IF;
90: (* B090 保持机械手抬升，D7 后退至 lrGripperBack；此时不是最终回位。 *)
aCommand[7] := F_Command(E_DeviceAction.Position, udiToken, stRecipe.lrGripperBack, stRecipe.lrPositionVelocity);
IF F_Done(aStatus[7], udiToken) THEN uiStep := 100; END_IF;
100: (* B100 后退到位后，G7 下降。 *)
aCommand[15] := F_Command(E_DeviceAction.Position, udiToken, 0.0, stRecipe.lrPositionVelocity);
IF F_Done(aStatus[15], udiToken) THEN uiStep := 110; END_IF;
110: (* B110 下降到位后，D7 再回 lrGripperHome；本支线结束前不允许送料。 *)
aCommand[7] := F_Command(E_DeviceAction.Position, udiToken, stRecipe.lrGripperHome, stRecipe.lrPositionVelocity);
IF F_Done(aStatus[7], udiToken) THEN uiStep := 1000; END_IF;
1000: (* 本支线完成，保持至 xExecute 撤销。 *) ;
ELSE xError := TRUE; udiErrorID := 4400;
END_CASE;
IF tonStep.Q THEN xError := TRUE; udiErrorID := 4400 + UINT_TO_UDINT(uiStep); END_IF;
END_IF;
xDone := xExecute AND (uiStep = 1000) AND NOT xError;

END_FUNCTION_BLOCK

// Device/Application/03_Units/FB_ReturnKnife
(* 模块说明：收尾支线 A：G5 喷油到设定时间，再令 D2 回刀。喷油仅在第一步保持请求。 *)
FUNCTION_BLOCK FB_ReturnKnife
VAR_INPUT
    xExecute : BOOL; (* 子流程执行许可；须保持到完成，清 FALSE 复位该流程步骤和错误。 *)
    stRecipe : ST_Recipe; (* 待校验配方或上层传入的运行配方，字段含义见 ST_Recipe。 *)
END_VAR
VAR_IN_OUT
    aCommand : ARRAY[1..17] OF ST_DeviceCommand; (* 统一设备请求数组 1..17；子流程写请求，设备管理器执行。 *)
    aStatus : ARRAY[1..17] OF ST_DeviceStatus; (* 各设备的反馈数组 1..17，供判断忙、完成序号、故障和位置。 *)
    udiCounter : UDINT; (* 全机共享的动作序号计数器，通过引用传递；由 F_NextID 分配，0 不使用。 *)
END_VAR
VAR_OUTPUT
    xDone : BOOL; (* 本子流程完成标志；执行许可撤销后复位。 *)
    xError : BOOL; (* 本设备或本子流程发生故障；具体原因见对应错误码。 *)
    udiErrorID : UDINT; (* 非法步骤码 4300；动作超时码=4300+uiStep，可据此定位本支线等待点。 *)
    uiStep : UINT; (* 当前子步骤：0 待机，10/20/... 执行动作，1000 完成；切勿在线强制跳步。 *)
END_VAR
VAR
    uiPrevStep : UINT := 65535; (* 上扫描步骤，用于判断本扫描是否刚进入新步骤。 *)
    udiToken : UDINT; (* 本步骤专用动作序号；同一步中的设备共用该号，以排除旧完成信号。 *)
    xEntry : BOOL; (* 本扫描为新步骤入口；用于分配新序号并复位步骤超时计时。 *)
    tonStep : TON; (* 步骤超时定时器；进入新步骤时复位，超时错误码由模块及当前步号组成。 *)
    tonSpray : TON; (* 通用子流程模板的喷油定时器，只有 FB_ReturnKnife 用其完成条件。 *)
END_VAR

(* 执行许可撤销即复位；步骤入口换新序号，每步等待本次动作完成，超时码=模块基码+步号。 *)
IF NOT xExecute THEN uiStep := 0; xError := FALSE; udiErrorID := 0; END_IF;
xEntry := uiStep <> uiPrevStep;
IF xEntry THEN udiToken := F_NextID(udiCounter); END_IF;
uiPrevStep := uiStep;
tonStep(IN := xExecute AND (uiStep > 0) AND (uiStep < 1000) AND NOT xEntry, PT := stRecipe.tStepTimeout);
tonSpray(IN := xExecute AND (uiStep = 10) AND aStatus[13].xActive, PT := stRecipe.tSpray);
IF xExecute AND NOT xError THEN
CASE uiStep OF
0: (* 待机；许可有效时进入首个动作。 *) uiStep := 10;
10: (* A010 G5 喷油并等待 tSpray；喷油建立后才开始计时。 *)
aCommand[13] := F_Command(E_DeviceAction.Run, udiToken, 0.0, 0.0);
IF tonSpray.Q THEN uiStep := 20; END_IF;
20: (* A020 结束喷油请求，D2 回到 lrCutHome，等待到位。 *)
aCommand[2] := F_Command(E_DeviceAction.Position, udiToken, stRecipe.lrCutHome, stRecipe.lrReturnVelocity);
IF F_Done(aStatus[2], udiToken) THEN uiStep := 1000; END_IF;
1000: (* 本支线完成，保持至 xExecute 撤销。 *) ;
ELSE xError := TRUE; udiErrorID := 4300;
END_CASE;
IF tonStep.Q THEN xError := TRUE; udiErrorID := 4300 + UINT_TO_UDINT(uiStep); END_IF;
END_IF;
xDone := xExecute AND (uiStep = 1000) AND NOT xError;

END_FUNCTION_BLOCK

// Device/Application/03_Units/FB_ClearanceUnit
(* 模块说明：并行执行 P/Q 两路避让；两路都完成才继续，任一路故障向主流程报告。 *)
FUNCTION_BLOCK FB_ClearanceUnit
VAR_INPUT
    xExecute : BOOL; (* 子流程执行许可；须保持到完成，清 FALSE 复位该流程步骤和错误。 *)
    stRecipe : ST_Recipe; (* 待校验配方或上层传入的运行配方，字段含义见 ST_Recipe。 *)
END_VAR
VAR_IN_OUT
    aCommand : ARRAY[1..17] OF ST_DeviceCommand; (* 统一设备请求数组 1..17；子流程写请求，设备管理器执行。 *)
    aStatus : ARRAY[1..17] OF ST_DeviceStatus; (* 各设备的反馈数组 1..17，供判断忙、完成序号、故障和位置。 *)
    udiCounter : UDINT; (* 全机共享的动作序号计数器，通过引用传递；由 F_NextID 分配，0 不使用。 *)
END_VAR
VAR_OUTPUT
    xDone : BOOL; (* 本子流程完成标志；执行许可撤销后复位。 *)
    xError : BOOL; (* 本设备或本子流程发生故障；具体原因见对应错误码。 *)
    udiErrorID : UDINT; (* 错误码；0 表示无错误，设备或流程发生异常时赋值。 *)
    uiLengthStep : UINT; (* 定长支线当前步骤，供监控定位等待点。 *)
    uiTransferStep : UINT; (* 流利条/侧推/侧挡支线当前步骤，供监控定位等待点。 *)
END_VAR
VAR
    fbLength : FB_ClearLength; (* P 支线：D5 升起、D4 移开。 *)
    fbTransfer : FB_ClearTransfer; (* 切割前流利条/侧推/侧挡避让支线。 *)
END_VAR

(* P/Q 两路同一扫描使能；xDone 使用 AND，任一路未完成均不得继续。 *)
fbLength(xExecute:=xExecute,stRecipe:=stRecipe,aCommand:=aCommand,aStatus:=aStatus,udiCounter:=udiCounter);
fbTransfer(xExecute:=xExecute,stRecipe:=stRecipe,aCommand:=aCommand,aStatus:=aStatus,udiCounter:=udiCounter);
xDone := fbLength.xDone AND fbTransfer.xDone;
xError := fbLength.xError OR fbTransfer.xError;
udiErrorID := MAX(fbLength.udiErrorID,fbTransfer.udiErrorID);
uiLengthStep := fbLength.uiStep; uiTransferStep := fbTransfer.uiStep;

END_FUNCTION_BLOCK

// Device/Application/03_Units/FB_ClearLength
(* 模块说明：切割前避让支线 P：D5 定长升起，再将 D4 移到避让位置。每步等待本次序号完成。 *)
FUNCTION_BLOCK FB_ClearLength
VAR_INPUT
    xExecute : BOOL; (* 子流程执行许可；须保持到完成，清 FALSE 复位该流程步骤和错误。 *)
    stRecipe : ST_Recipe; (* 待校验配方或上层传入的运行配方，字段含义见 ST_Recipe。 *)
END_VAR
VAR_IN_OUT
    aCommand : ARRAY[1..17] OF ST_DeviceCommand; (* 统一设备请求数组 1..17；子流程写请求，设备管理器执行。 *)
    aStatus : ARRAY[1..17] OF ST_DeviceStatus; (* 各设备的反馈数组 1..17，供判断忙、完成序号、故障和位置。 *)
    udiCounter : UDINT; (* 全机共享的动作序号计数器，通过引用传递；由 F_NextID 分配，0 不使用。 *)
END_VAR
VAR_OUTPUT
    xDone : BOOL; (* 本子流程完成标志；执行许可撤销后复位。 *)
    xError : BOOL; (* 本设备或本子流程发生故障；具体原因见对应错误码。 *)
    udiErrorID : UDINT; (* 非法步骤码 4100；动作超时码=4100+uiStep，可据此定位本支线等待点。 *)
    uiStep : UINT; (* 当前子步骤：0 待机，10/20/... 执行动作，1000 完成；切勿在线强制跳步。 *)
END_VAR
VAR
    uiPrevStep : UINT := 65535; (* 上扫描步骤，用于判断本扫描是否刚进入新步骤。 *)
    udiToken : UDINT; (* 本步骤专用动作序号；同一步中的设备共用该号，以排除旧完成信号。 *)
    xEntry : BOOL; (* 本扫描为新步骤入口；用于分配新序号并复位步骤超时计时。 *)
    tonStep : TON; (* 步骤超时定时器；进入新步骤时复位，超时错误码由模块及当前步号组成。 *)
    tonSpray : TON; (* 通用子流程模板的喷油定时器，只有 FB_ReturnKnife 用其完成条件。 *)
END_VAR

(* 执行许可撤销即复位；步骤入口换新序号，每步等待本次动作完成，超时码=模块基码+步号。 *)
IF NOT xExecute THEN uiStep := 0; xError := FALSE; udiErrorID := 0; END_IF;
xEntry := uiStep <> uiPrevStep;
IF xEntry THEN udiToken := F_NextID(udiCounter); END_IF;
uiPrevStep := uiStep;
tonStep(IN := xExecute AND (uiStep > 0) AND (uiStep < 1000) AND NOT xEntry, PT := stRecipe.tStepTimeout);
tonSpray(IN := xExecute AND (uiStep = 10) AND aStatus[13].xActive, PT := stRecipe.tSpray);
IF xExecute AND NOT xError THEN
CASE uiStep OF
0: (* 待机；许可有效时进入首个动作。 *) uiStep := 10;
10: (* P010 定长 D5 升起避让；确认本次动作完成后再允许 D4 平移。 *)
aCommand[5] := F_Command(E_DeviceAction.Position, udiToken, 0.0, stRecipe.lrPositionVelocity);
IF F_Done(aStatus[5], udiToken) THEN uiStep := 20; END_IF;
20: (* P020 定长 D4 移到配方避让位置，等待本次序号完成。 *)
aCommand[4] := F_Command(E_DeviceAction.Position, udiToken, stRecipe.lrLengthClear, stRecipe.lrPositionVelocity);
IF F_Done(aStatus[4], udiToken) THEN uiStep := 1000; END_IF;
1000: (* 本支线完成，保持至 xExecute 撤销。 *) ;
ELSE xError := TRUE; udiErrorID := 4100;
END_CASE;
IF tonStep.Q THEN xError := TRUE; udiErrorID := 4100 + UINT_TO_UDINT(uiStep); END_IF;
END_IF;
xDone := xExecute AND (uiStep = 1000) AND NOT xError;

END_FUNCTION_BLOCK

// Device/Application/03_Units/FB_ClearTransfer
(* 模块说明：切割前避让支线 Q：G4 流利条下降、G3 解除侧推、G2 侧挡下降。 *)
FUNCTION_BLOCK FB_ClearTransfer
VAR_INPUT
    xExecute : BOOL; (* 子流程执行许可；须保持到完成，清 FALSE 复位该流程步骤和错误。 *)
    stRecipe : ST_Recipe; (* 待校验配方或上层传入的运行配方，字段含义见 ST_Recipe。 *)
END_VAR
VAR_IN_OUT
    aCommand : ARRAY[1..17] OF ST_DeviceCommand; (* 统一设备请求数组 1..17；子流程写请求，设备管理器执行。 *)
    aStatus : ARRAY[1..17] OF ST_DeviceStatus; (* 各设备的反馈数组 1..17，供判断忙、完成序号、故障和位置。 *)
    udiCounter : UDINT; (* 全机共享的动作序号计数器，通过引用传递；由 F_NextID 分配，0 不使用。 *)
END_VAR
VAR_OUTPUT
    xDone : BOOL; (* 本子流程完成标志；执行许可撤销后复位。 *)
    xError : BOOL; (* 本设备或本子流程发生故障；具体原因见对应错误码。 *)
    udiErrorID : UDINT; (* 非法步骤码 4200；动作超时码=4200+uiStep，可据此定位本支线等待点。 *)
    uiStep : UINT; (* 当前子步骤：0 待机，10/20/... 执行动作，1000 完成；切勿在线强制跳步。 *)
END_VAR
VAR
    uiPrevStep : UINT := 65535; (* 上扫描步骤，用于判断本扫描是否刚进入新步骤。 *)
    udiToken : UDINT; (* 本步骤专用动作序号；同一步中的设备共用该号，以排除旧完成信号。 *)
    xEntry : BOOL; (* 本扫描为新步骤入口；用于分配新序号并复位步骤超时计时。 *)
    tonStep : TON; (* 步骤超时定时器；进入新步骤时复位，超时错误码由模块及当前步号组成。 *)
    tonSpray : TON; (* 通用子流程模板的喷油定时器，只有 FB_ReturnKnife 用其完成条件。 *)
END_VAR

(* 执行许可撤销即复位；步骤入口换新序号，每步等待本次动作完成，超时码=模块基码+步号。 *)
IF NOT xExecute THEN uiStep := 0; xError := FALSE; udiErrorID := 0; END_IF;
xEntry := uiStep <> uiPrevStep;
IF xEntry THEN udiToken := F_NextID(udiCounter); END_IF;
uiPrevStep := uiStep;
tonStep(IN := xExecute AND (uiStep > 0) AND (uiStep < 1000) AND NOT xEntry, PT := stRecipe.tStepTimeout);
tonSpray(IN := xExecute AND (uiStep = 10) AND aStatus[13].xActive, PT := stRecipe.tSpray);
IF xExecute AND NOT xError THEN
CASE uiStep OF
0: (* 待机；许可有效时进入首个动作。 *) uiStep := 10;
10: (* Q010 流利条 G4 下降。 *)
aCommand[12] := F_Command(E_DeviceAction.Position, udiToken, 0.0, stRecipe.lrPositionVelocity);
IF F_Done(aStatus[12], udiToken) THEN uiStep := 20; END_IF;
20: (* Q020 推动气缸 G3 放开。 *)
aCommand[11] := F_Command(E_DeviceAction.Position, udiToken, 0.0, stRecipe.lrPositionVelocity);
IF F_Done(aStatus[11], udiToken) THEN uiStep := 30; END_IF;
30: (* Q030 侧挡 G2 下降。目标固定发 1.0：本层不知道侧挡是单缸还是 300/450/600 三缸组，
   由设备层自己解释——仿真气缸按 1.0 到伸出端，真实三缸组按当前料型选缸下降。 *)
aCommand[10] := F_Command(E_DeviceAction.Position, udiToken, 1.0, stRecipe.lrPositionVelocity);
IF F_Done(aStatus[10], udiToken) THEN uiStep := 1000; END_IF;
1000: (* 本支线完成，保持至 xExecute 撤销。 *) ;
ELSE xError := TRUE; udiErrorID := 4200;
END_CASE;
IF tonStep.Q THEN xError := TRUE; udiErrorID := 4200 + UINT_TO_UDINT(uiStep); END_IF;
END_IF;
xDone := xExecute AND (uiStep = 1000) AND NOT xError;

END_FUNCTION_BLOCK

// Device/Application/03_Units/FB_PostCut
(* 模块说明：切割后先 G9 抬刀，再 G1 抬压；之后同时执行回刀、机械手移料、定长复位，三路全完成才结束。 *)
FUNCTION_BLOCK FB_PostCut
VAR_INPUT
    xExecute : BOOL; (* 子流程执行许可；须保持到完成，清 FALSE 复位该流程步骤和错误。 *)
    stRecipe : ST_Recipe; (* 待校验配方或上层传入的运行配方，字段含义见 ST_Recipe。 *)
END_VAR
VAR_IN_OUT
    aCommand : ARRAY[1..17] OF ST_DeviceCommand; (* 统一设备请求数组 1..17；子流程写请求，设备管理器执行。 *)
    aStatus : ARRAY[1..17] OF ST_DeviceStatus; (* 各设备的反馈数组 1..17，供判断忙、完成序号、故障和位置。 *)
    udiCounter : UDINT; (* 全机共享的动作序号计数器，通过引用传递；由 F_NextID 分配，0 不使用。 *)
END_VAR
VAR_OUTPUT
    xDone : BOOL; (* 本子流程完成标志；执行许可撤销后复位。 *)
    xError : BOOL; (* 本设备或本子流程发生故障；具体原因见对应错误码。 *)
    udiErrorID : UDINT; (* 非法总步骤为 4700，超时为 4700+总步号；支线故障则向上传递支线错误码。 *)
    uiStep : UINT; (* 当前子步骤：0 待机，10/20/... 执行动作，1000 完成；切勿在线强制跳步。 *)
    uiKnifeStep : UINT; (* 收尾回刀支线 A 当前步骤：喷油、回刀或完成。 *)
    uiUnloadStep : UINT; (* 机械手移料支线 B 步骤，10..110 每步加 10，1000 完成；详见 FB_Unload。 *)
    uiLengthStep : UINT; (* 定长支线当前步骤，供监控定位等待点。 *)
END_VAR
VAR
    fbKnife : FB_ReturnKnife; (* 收尾支线 A：喷油后回刀。 *)
    fbUnload : FB_Unload; (* 收尾支线 B：机械手移料，含后退、下降、最终回位。 *)
    fbLength : FB_ResetLength; (* C 支线：D4 回检测位置、D5 下降、确认下降到位。 *)
    uiPrevStep : UINT := 65535; (* 上扫描步骤，用于判断本扫描是否刚进入新步骤。 *)
    udiToken : UDINT; (* 本步骤专用动作序号；同一步中的设备共用该号，以排除旧完成信号。 *)
    xEntry : BOOL; (* 本扫描为新步骤入口；用于分配新序号并复位步骤超时计时。 *)
    tonStep : TON; (* 步骤超时定时器；进入新步骤时复位，超时错误码由模块及当前步号组成。 *)
END_VAR

IF NOT xExecute THEN uiStep := 0; xError := FALSE; udiErrorID := 0; END_IF
(* 每个总步骤分配新序号；等待三路期间保留总步骤超时。 *)
xEntry := uiStep <> uiPrevStep;
IF xEntry THEN udiToken := F_NextID(udiCounter); END_IF
uiPrevStep := uiStep;
tonStep(IN:=xExecute AND NOT xEntry AND (uiStep>0) AND (uiStep<1000),PT:=stRecipe.tStepTimeout);
IF xExecute AND NOT xError THEN
    CASE uiStep OF
    0: (* 待机，执行许可有效后进入抬刀。 *) uiStep := 10;
    10: (* 先 G9 盘刀提升；同时保持 G1 下压，刀没抬起来之前不能松压板。 *)
        aCommand[9] := F_Command(E_DeviceAction.Position,udiToken,1.0,stRecipe.lrPositionVelocity);
        aCommand[17] := F_Command(E_DeviceAction.Position,udiToken,0.0,stRecipe.lrPositionVelocity);
        IF F_Done(aStatus[17],udiToken) THEN uiStep := 20; END_IF
    20: (* 再 G1 下压提升，等待本次序号完成。 *)
        aCommand[9] := F_Command(E_DeviceAction.Position,udiToken,0.0,stRecipe.lrPositionVelocity);
        IF F_Done(aStatus[9],udiToken) THEN uiStep := 30; END_IF
    30: (* 等待回刀、机械手移料、定长复位三路全部完成。 *)
        IF fbKnife.xDone AND fbUnload.xDone AND fbLength.xDone THEN uiStep := 1000; END_IF
    1000: (* 三路收尾结束，保持完成反馈直到执行许可撤销。 *) ;
    ELSE xError := TRUE; udiErrorID := 4700;
    END_CASE
    IF tonStep.Q THEN xError := TRUE; udiErrorID := 4700+UINT_TO_UDINT(uiStep); END_IF
END_IF
(* 三路只在总步骤 30 同时使能，并且每扫描调用；等待三路全完成才退出。 *)
fbKnife(xExecute:=xExecute AND (uiStep=30),stRecipe:=stRecipe,aCommand:=aCommand,aStatus:=aStatus,udiCounter:=udiCounter);
fbUnload(xExecute:=xExecute AND (uiStep=30),stRecipe:=stRecipe,aCommand:=aCommand,aStatus:=aStatus,udiCounter:=udiCounter);
fbLength(xExecute:=xExecute AND (uiStep=30),stRecipe:=stRecipe,aCommand:=aCommand,aStatus:=aStatus,udiCounter:=udiCounter);
IF fbKnife.xError OR fbUnload.xError OR fbLength.xError THEN
    xError:=TRUE; udiErrorID:=MAX(fbKnife.udiErrorID,MAX(fbUnload.udiErrorID,fbLength.udiErrorID));
END_IF
xDone := xExecute AND (uiStep=1000) AND NOT xError;
uiKnifeStep:=fbKnife.uiStep; uiUnloadStep:=fbUnload.uiStep; uiLengthStep:=fbLength.uiStep;

END_FUNCTION_BLOCK

// Device/Application/03_Units/FB_ResetLength
(* 模块说明：收尾支线 C：D4 回检测位置、D5 下降到位、确认下降位置；随后具备来料检测条件。 *)
FUNCTION_BLOCK FB_ResetLength
VAR_INPUT
    xExecute : BOOL; (* 子流程执行许可；须保持到完成，清 FALSE 复位该流程步骤和错误。 *)
    stRecipe : ST_Recipe; (* 待校验配方或上层传入的运行配方，字段含义见 ST_Recipe。 *)
END_VAR
VAR_IN_OUT
    aCommand : ARRAY[1..17] OF ST_DeviceCommand; (* 统一设备请求数组 1..17；子流程写请求，设备管理器执行。 *)
    aStatus : ARRAY[1..17] OF ST_DeviceStatus; (* 各设备的反馈数组 1..17，供判断忙、完成序号、故障和位置。 *)
    udiCounter : UDINT; (* 全机共享的动作序号计数器，通过引用传递；由 F_NextID 分配，0 不使用。 *)
END_VAR
VAR_OUTPUT
    xDone : BOOL; (* 本子流程完成标志；执行许可撤销后复位。 *)
    xError : BOOL; (* 本设备或本子流程发生故障；具体原因见对应错误码。 *)
    udiErrorID : UDINT; (* 非法步骤码 4500；动作超时码=4500+uiStep，可据此定位本支线等待点。 *)
    uiStep : UINT; (* 当前子步骤：0 待机，10/20/... 执行动作，1000 完成；切勿在线强制跳步。 *)
END_VAR
VAR
    uiPrevStep : UINT := 65535; (* 上扫描步骤，用于判断本扫描是否刚进入新步骤。 *)
    udiToken : UDINT; (* 本步骤专用动作序号；同一步中的设备共用该号，以排除旧完成信号。 *)
    xEntry : BOOL; (* 本扫描为新步骤入口；用于分配新序号并复位步骤超时计时。 *)
    tonStep : TON; (* 步骤超时定时器；进入新步骤时复位，超时错误码由模块及当前步号组成。 *)
    tonSpray : TON; (* 通用子流程模板的喷油定时器，只有 FB_ReturnKnife 用其完成条件。 *)
END_VAR

(* 执行许可撤销即复位；步骤入口换新序号，每步等待本次动作完成，超时码=模块基码+步号。 *)
IF NOT xExecute THEN uiStep := 0; xError := FALSE; udiErrorID := 0; END_IF;
xEntry := uiStep <> uiPrevStep;
IF xEntry THEN udiToken := F_NextID(udiCounter); END_IF;
uiPrevStep := uiStep;
tonStep(IN := xExecute AND (uiStep > 0) AND (uiStep < 1000) AND NOT xEntry, PT := stRecipe.tStepTimeout);
tonSpray(IN := xExecute AND (uiStep = 10) AND aStatus[13].xActive, PT := stRecipe.tSpray);
IF xExecute AND NOT xError THEN
CASE uiStep OF
0: (* 待机；许可有效时进入首个动作。 *) uiStep := 10;
10: (* C010 定长 D4 回到配方检测位置 lrLengthPosition。 *)
aCommand[4] := F_Command(E_DeviceAction.Position, udiToken, stRecipe.lrLengthPosition, stRecipe.lrPositionVelocity);
IF F_Done(aStatus[4], udiToken) THEN uiStep := 20; END_IF;
20: (* C020 D4 到位后，定长 D5 下降。 *)
aCommand[5] := F_Command(E_DeviceAction.Position, udiToken, 1.0, stRecipe.lrPositionVelocity);
IF F_Done(aStatus[5], udiToken) THEN uiStep := 30; END_IF;
30: (* C030 确认 D5 下降端到位，后续送料才具备光电检测条件。 *)
IF F_At(aStatus[5],1.0) THEN uiStep := 1000; END_IF;
1000: (* 本支线完成，保持至 xExecute 撤销。 *) ;
ELSE xError := TRUE; udiErrorID := 4500;
END_CASE;
IF tonStep.Q THEN xError := TRUE; udiErrorID := 4500 + UINT_TO_UDINT(uiStep); END_IF;
END_IF;
xDone := xExecute AND (uiStep = 1000) AND NOT xError;

END_FUNCTION_BLOCK

// Device/Application/03_Units/FB_Initialize
(* 模块说明：初始姿态整理流程。20 步摆好避让姿态后，25 步让真实轴回零，30 步再按配方绝对定位。 *)
FUNCTION_BLOCK FB_Initialize
VAR_INPUT
    xExecute : BOOL; (* 子流程执行许可；须保持到完成，清 FALSE 复位该流程步骤和错误。 *)
    stRecipe : ST_Recipe; (* 待校验配方或上层传入的运行配方，字段含义见 ST_Recipe。 *)
END_VAR
VAR_IN_OUT
    aCommand : ARRAY[1..17] OF ST_DeviceCommand; (* 统一设备请求数组 1..17；子流程写请求，设备管理器执行。 *)
    aStatus : ARRAY[1..17] OF ST_DeviceStatus; (* 各设备的反馈数组 1..17，供判断忙、完成序号、故障和位置。 *)
    udiCounter : UDINT; (* 全机共享的动作序号计数器，通过引用传递；由 F_NextID 分配，0 不使用。 *)
END_VAR
VAR_OUTPUT
    xDone : BOOL; (* 本子流程完成标志；执行许可撤销后复位。 *)
    xError : BOOL; (* 本设备或本子流程发生故障；具体原因见对应错误码。 *)
    udiErrorID : UDINT; (* 非法步骤码 4600；动作超时码=4600+uiStep，可据此定位本支线等待点。 *)
    uiStep : UINT; (* 当前子步骤：0 待机，10/20/25/30/40 执行动作，1000 完成；切勿在线强制跳步。 *)
END_VAR
VAR
    uiPrevStep : UINT := 65535; (* 上扫描步骤，用于判断本扫描是否刚进入新步骤。 *)
    udiToken : UDINT; (* 本步骤专用动作序号；同一步中的设备共用该号，以排除旧完成信号。 *)
    xEntry : BOOL; (* 本扫描为新步骤入口；用于分配新序号并复位步骤超时计时。 *)
    tonStep : TON; (* 步骤超时定时器；进入新步骤时复位，超时错误码由模块及当前步号组成。 *)
    tonSpray : TON; (* 通用子流程模板的喷油定时器，只有 FB_ReturnKnife 用其完成条件。 *)
END_VAR

(* 执行许可撤销即复位；步骤入口换新序号，每步等待本次动作完成，超时码=模块基码+步号。 *)
IF NOT xExecute THEN uiStep := 0; xError := FALSE; udiErrorID := 0; END_IF;
xEntry := uiStep <> uiPrevStep;
IF xEntry THEN udiToken := F_NextID(udiCounter); END_IF;
uiPrevStep := uiStep;
tonStep(IN := xExecute AND (uiStep > 0) AND (uiStep < 1000) AND NOT xEntry, PT := stRecipe.tStepTimeout);
tonSpray(IN := xExecute AND (uiStep = 10) AND aStatus[13].xActive, PT := stRecipe.tSpray);
IF xExecute AND NOT xError THEN
CASE uiStep OF
0: (* 待机；许可有效时进入首个动作。 *) uiStep := 10;
10: (* 仿真初始化 10：同时抬起 G9、抬起 G1、打开 G8，三项都完成才继续。 *)
aCommand[17] := F_Command(E_DeviceAction.Position, udiToken, 0.0, stRecipe.lrPositionVelocity);
aCommand[9] := F_Command(E_DeviceAction.Position, udiToken, 0.0, stRecipe.lrPositionVelocity);
aCommand[16] := F_Command(E_DeviceAction.Position, udiToken, 0.0, stRecipe.lrPositionVelocity);
IF F_Done(aStatus[17], udiToken) AND F_Done(aStatus[9], udiToken) AND F_Done(aStatus[16], udiToken) THEN uiStep := 20; END_IF;
20: (* 仿真初始化 20：D5 升起、G2 提升、G3 释放、G4 提升、G7 下降，全部完成再定位。 *)
aCommand[5] := F_Command(E_DeviceAction.Position, udiToken, 0.0, stRecipe.lrPositionVelocity);
aCommand[10] := F_Command(E_DeviceAction.Position, udiToken, 0.0, stRecipe.lrPositionVelocity);
aCommand[11] := F_Command(E_DeviceAction.Position, udiToken, 0.0, stRecipe.lrPositionVelocity);
aCommand[12] := F_Command(E_DeviceAction.Position, udiToken, 1.0, stRecipe.lrPositionVelocity);
aCommand[15] := F_Command(E_DeviceAction.Position, udiToken, 0.0, stRecipe.lrPositionVelocity);
IF F_Done(aStatus[5], udiToken) AND F_Done(aStatus[10], udiToken) AND F_Done(aStatus[11], udiToken) AND F_Done(aStatus[12], udiToken) AND F_Done(aStatus[15], udiToken) THEN uiStep := 25; END_IF;
25: (* 初始化 25：真实轴回零。D2 走刀与 D8 旋转是真轴，D4 定长平移当前为仿真，由仿真在 tSimAction 后完成。
       D3 盘刀是连续旋转主轴，自动流程只下发 Run 不定位，因此不参与回零，也不占本步完成条件。 *)
aCommand[2] := F_Command(E_DeviceAction.Home, udiToken, 0.0, 0.0);
aCommand[4] := F_Command(E_DeviceAction.Home, udiToken, 0.0, 0.0);
aCommand[8] := F_Command(E_DeviceAction.Home, udiToken, 0.0, 0.0);
IF F_Done(aStatus[2], udiToken) AND F_Done(aStatus[4], udiToken) AND F_Done(aStatus[8], udiToken) THEN uiStep := 30; END_IF;
30: (* 仿真初始化 30：D2/D4/D7/D8 移至示例初始坐标，全部完成才继续。 *)
aCommand[2] := F_Command(E_DeviceAction.Position, udiToken, stRecipe.lrCutHome, stRecipe.lrPositionVelocity);
aCommand[4] := F_Command(E_DeviceAction.Position, udiToken, stRecipe.lrLengthPosition, stRecipe.lrPositionVelocity);
aCommand[7] := F_Command(E_DeviceAction.Position, udiToken, stRecipe.lrGripperHome, stRecipe.lrPositionVelocity);
aCommand[8] := F_Command(E_DeviceAction.Position, udiToken, 0.0, stRecipe.lrPositionVelocity);
IF F_Done(aStatus[2], udiToken) AND F_Done(aStatus[4], udiToken) AND F_Done(aStatus[7], udiToken) AND F_Done(aStatus[8], udiToken) THEN uiStep := 40; END_IF;
40: (* 仿真初始化 40：D5 下降，准备进入来料检测。 *)
aCommand[5] := F_Command(E_DeviceAction.Position, udiToken, 1.0, stRecipe.lrPositionVelocity);
IF F_Done(aStatus[5], udiToken) THEN uiStep := 1000; END_IF;
1000: (* 本支线完成，保持至 xExecute 撤销。 *) ;
ELSE xError := TRUE; udiErrorID := 4600;
END_CASE;
IF tonStep.Q THEN xError := TRUE; udiErrorID := 4600 + UINT_TO_UDINT(uiStep); END_IF;
END_IF;
xDone := xExecute AND (uiStep = 1000) AND NOT xError;

END_FUNCTION_BLOCK

// Device/Application/04_Machine/FB_Interlocks
(* 模块说明：对手动、初始化和自动请求统一执行软件互锁。禁止动作时改为停止，并报告最后一个被阻挡设备。 *)
FUNCTION_BLOCK FB_Interlocks
VAR_INPUT
	xPermit : BOOL; (* 整机当前允许发出动作的总许可；仍需继续满足各设备互锁。 *)
	xManualMode : BOOL; (* 当前处于手动模式；手动模式暂不做机构互锁，互锁只约束自动流程。 *)
	stRecipe : ST_Recipe; (* 待校验配方或上层传入的运行配方，字段含义见 ST_Recipe。 *)
	stReal : ST_RealDeviceSettings; (* 真实设备接管设置；预留输入，当前手动已默认不查互锁，判定未使用。 *)
    tViolationDelay : TIME := T#200MS; (* 机构违规确认时间；连续保持这么久才认定，避免过渡瞬间误报。 *)
	aRequest : ARRAY[1..17] OF ST_DeviceCommand; (* 初始化/手动/自动产生的原始请求，每周期先清空，再交互锁筛选。 *)
	aStatus : ARRAY[1..17] OF ST_DeviceStatus; (* 各设备的反馈数组 1..17，供判断忙、完成序号、故障和位置。 *)
END_VAR
VAR_OUTPUT
	aCommand : ARRAY[1..17] OF ST_DeviceCommand; (* 统一设备请求数组 1..17；子流程写请求，设备管理器执行。 *)
	uiBlockedDevice : UINT; (* 本扫描最后一个被互锁阻挡的设备索引；0 表示无阻挡，可结合设备状态排查。 *)
    xViolated : BOOL; (* 机构互锁违规已确认：总许可通过、但机构条件不满足，且持续超过确认时间。 *)
    uiViolatedDevice : UINT; (* 确认违规的设备索引；0 表示无。 *)
END_VAR
VAR
	i : INT; (* 本扫描数组遍历索引；含义及范围以当前 FOR 循环为准。 *)
	xAllowed : BOOL; (* 当前遍历设备的最终互锁允许结果。 *)
	xMotion : BOOL; (* 当前请求是否为点动或离开当前位置的定位，决定是否检查机构避让。 *)
	xKnifeUp : BOOL; (* G9 刀具处于提升端且设备无忙无故障。 *)
	xPressUp : BOOL; (* G1 下压机构处于抬起端且设备无忙无故障。 *)
	xClampOpen : BOOL; (* G8 夹爪处于打开端且设备无忙无故障。 *)
    xPermitOK : BOOL; (* 仅总许可结果；用来区分"许可没通过"和"机构条件不满足"。 *)
    xStructBlocked : BOOL; (* 本扫描是否有请求因机构条件被拒。 *)
    uiStructDevice : UINT; (* 最后一个因机构条件被拒的设备索引。 *)
    tonViolation : TON; (* 机构违规去抖定时器。 *)
END_VAR

(* 以下为普通程序互锁；实际急停、门锁、失气等安全功能须由最终硬件方案实现。 *)
uiBlockedDevice:=0;
    xStructBlocked:=FALSE;
    uiStructDevice:=UINT#0;
xKnifeUp:=F_At(aStatus[17],0.0); xPressUp:=F_At(aStatus[9],0.0);
xClampOpen:=F_At(aStatus[16],0.0);
FOR i:=1 TO 17 DO
    aCommand[i]:=aRequest[i];
    xPermitOK:=xPermit AND (i<>6);
    xAllowed:=xPermitOK;
    xMotion:=(aRequest[i].eAction=E_DeviceAction.Jog) OR
        ((aRequest[i].eAction=E_DeviceAction.Position) AND
        (ABS(aRequest[i].lrTarget-aStatus[i].lrPosition)>0.01));
    (* 手动模式暂不做机构互锁：单轴调试要求能独立动作，互锁只约束自动流程。
       手动下的硬干涉（D5 挡 D4 行程、平台旋转扫刀等）后续按调试情况逐条补回。
       xPermit 不受此影响，任何时候都要先满足。 *)
    IF xMotion AND NOT xManualMode THEN
        CASE i OF
        (* D4 平移之前，D5 定长升降必须已经升起。 *)
        4: xAllowed:=xAllowed AND F_At(aStatus[5],0.0);
        (* D8 平台旋转之前，盘刀和下压抬起、G3 侧推解除。 *)
        8: xAllowed:=xAllowed AND xKnifeUp AND xPressUp AND F_At(aStatus[11],0.0);
        (* G1 下压时，平台不得旋转，盘刀抬起且 D2 在回刀起点。 *)
        9:
            IF aRequest[i].lrTarget>0.5 THEN
                xAllowed:=xAllowed AND NOT aStatus[8].xBusy AND xKnifeUp AND F_At(aStatus[2],stRecipe.lrCutHome);
            ELSE
                (* 抬起前盘刀必须先抬起，否则刀还在工件里就松了压板。 *)
                xAllowed:=xAllowed AND xKnifeUp;
            END_IF
        (* G9 下刀时，下压到位、旋转停止、定长升起、流利条下降、侧挡下降。 *)
        17:
            IF aRequest[i].lrTarget>0.5 THEN
                xAllowed:=xAllowed AND F_At(aStatus[9],1.0) AND NOT aStatus[8].xBusy
                    AND F_At(aStatus[5],0.0) AND F_At(aStatus[12],0.0) AND F_At(aStatus[10],1.0);
            END_IF
        (* D2 正向切割需下压和盘刀下降到位且盘刀运行；回刀需盘刀抬起。 *)
        2:
            IF ((aRequest[i].eAction=E_DeviceAction.Position) AND (aRequest[i].lrTarget>stRecipe.lrCutHome+0.01))
               OR ((aRequest[i].eAction=E_DeviceAction.Jog) AND (aRequest[i].lrVelocity>0.0)) THEN
                xAllowed:=xAllowed AND F_At(aStatus[9],1.0) AND F_At(aStatus[17],1.0) AND aStatus[3].xActive;
            ELSE xAllowed:=xAllowed AND xKnifeUp;
            END_IF
        (* D7 机械手分点动、拉料、抬升平移与下降回位分别校验，保持后退/下降/回位顺序。 *)
        7:
            xAllowed:=xAllowed AND xKnifeUp AND xPressUp;
            IF aRequest[i].eAction=E_DeviceAction.Jog THEN
                xAllowed:=xAllowed AND F_At(aStatus[15],1.0) AND xClampOpen;
            ELSIF ABS(aRequest[i].lrTarget-stRecipe.lrGripperHome)<0.01 THEN
                xAllowed:=xAllowed AND F_At(aStatus[15],0.0) AND xClampOpen;
            ELSIF ABS(aRequest[i].lrTarget-stRecipe.lrGripperPull)<0.01 THEN
                xAllowed:=xAllowed AND F_At(aStatus[15],1.0) AND F_At(aStatus[16],1.0);
            ELSE xAllowed:=xAllowed AND F_At(aStatus[15],1.0) AND xClampOpen;
            END_IF
        END_CASE
    END_IF
    (* 互锁不满足则用 Stop 覆盖该设备请求；记录最后一个被阻挡编号，便于排查。 *)
    IF NOT xAllowed THEN
        IF aRequest[i].eAction<>E_DeviceAction.None THEN
            uiBlockedDevice:=INT_TO_UINT(i);
            (* 只有总许可通过时的拒绝才算机构违规；许可未通过已由 1001 等上报，不在这里重复。 *)
            IF xPermitOK THEN
                xStructBlocked:=TRUE;
                uiStructDevice:=INT_TO_UINT(i);
            END_IF
        END_IF
        aCommand[i].eAction:=E_DeviceAction.Stop;
    END_IF
END_FOR
tonViolation(IN:=xStructBlocked,PT:=tViolationDelay);
xViolated:=tonViolation.Q;
IF xViolated THEN uiViolatedDevice:=uiStructDevice; ELSE uiViolatedDevice:=UINT#0; END_IF

END_FUNCTION_BLOCK

// Device/Application/04_Machine/FB_AlarmManager
(* 模块说明：锁存首次非零报警。只有复位有效且当前没有新报警时清除；同一扫描有新报警时仍会锁存。 *)
FUNCTION_BLOCK FB_AlarmManager
VAR_INPUT
    udiIncoming : UDINT; (* 当前扫描的新报警码；0 表示当前未提出报警。 *)
    xReset : BOOL; (* 故障复位许可；仿真设备仅在故障注入已撤销时清除错误。 *)
END_VAR
VAR_OUTPUT
    udiLatched : UDINT; (* 已锁存的首个非零报警码；后续报警不覆盖，满足复位条件后清零。 *)
END_VAR

(* 只有没有当前报警原因才清锁存；当前代码保留第一个非零报警，后续报警不覆盖。 *)
IF xReset AND (udiIncoming=0) THEN udiLatched:=0; END_IF
IF (udiLatched=0) AND (udiIncoming<>0) THEN udiLatched:=udiIncoming; END_IF

END_FUNCTION_BLOCK

// Device/Application/02_Devices/F_SafetyBypassActive
(* 模块说明：安全许可软件旁路的唯一判定点。两级开关同时置位才返回 TRUE。 *)
FUNCTION F_SafetyBypassActive : BOOL
VAR_IN_OUT
	stReal : ST_RealDeviceSettings; (* 引用传递，避免每次扫描拷贝整个设置结构体。 *)
END_VAR

(* 一级开关与二级确认必须同时置位；任一为 FALSE 就返回 FALSE，保持原有安全逻辑。 *)
F_SafetyBypassActive := stReal.xSafetyBypass AND stReal.xSafetyBypassConfirm;

END_FUNCTION

// Device/Application/04_Machine/FB_PanelInput
(* 模块说明：每扫描先读取实体面板或仿真面板，形成唯一的本地命令来源。上位机不能修改此处的模式。 *)
FUNCTION_BLOCK FB_PanelInput
VAR_INPUT
    xSimulation : BOOL; (* TRUE 使用内部仿真；当前 FALSE 报未实现 3001，不会接管真实运动。 *)
    stReal : ST_PanelInputs; (* 从物理 I/O 映射得到的标准化面板输入，当前未分配端子地址。 *)
    stSim : ST_PanelInputs; (* 仿真用面板输入，代替尚未连接的实体旋钮和按钮。 *)
    xContinuous : BOOL; (* TRUE 连续循环；FALSE 在当前完整循环结束后回到就绪。 *)
    xUseRealPanel : BOOL := TRUE; (* TRUE 取实体面板 stReal；FALSE 取仿真面板 stSim。与 xSimulation 解耦，后者恒为 TRUE。 *)
END_VAR
VAR_OUTPUT
    stCommand : ST_OperatorCommand; (* 由本地面板生成的命令，模式仅由 xAutoMode 形成。 *)
END_VAR
VAR
    stSelected : ST_PanelInputs; (* 本扫描选中的实体/仿真面板输入快照。 *)
END_VAR

(* 这里只处理已归一化的逻辑信号；端子、常开/常闭和必要的输入滤波在实际 I/O 映射时确定。
   面板来源与 xSimulation 解耦：设备可以全仿真而面板用实物按钮，也可以反过来。 *)
IF xUseRealPanel THEN stSelected:=stReal;
ELSE stSelected:=stSim; END_IF
(* 默认手动，只有本地旋钮明确选择自动才转自动；急停反馈不混入普通停止按钮。 *)
stCommand.eMode:=E_MachineMode.Manual;
IF stSelected.xAutoMode THEN stCommand.eMode:=E_MachineMode.Automatic; END_IF
stCommand.xInitialize:=stSelected.xInitialize;
stCommand.xStart:=stSelected.xStart;
stCommand.xStop:=stSelected.xStop;
stCommand.xResetAlarm:=stSelected.xResetAlarm;
stCommand.xContinuous:=xContinuous;
(* 启动/停止是"按一下切换"的两个独立按钮，这里只做电平搬运；
   沿检测与运行态锁存放在 FB_Machine，保证停机判据全机只有一处。 *)
stCommand.xRunStart:=stSelected.xRunStart;
stCommand.xRunStop:=stSelected.xRunStop;

END_FUNCTION_BLOCK

// Device/Application/05_Communication/FB_ModbusInterface
(* 模块说明：Modbus 协议 v2：只解析可选的远程启动/停止，发布整机状态。模式只读；参数映射另行配置。 *)
FUNCTION_BLOCK FB_ModbusInterface
VAR_INPUT
    xEnable : BOOL; (* 通信解析许可；首次使能只记录现有序号，防止重放旧命令。 *)
    stStatus : ST_MachineStatus; (* 本模块对外发布的状态；字段含义见其数据类型。 *)
    aStatus : ARRAY[1..17] OF ST_DeviceStatus; (* 各设备的反馈数组 1..17，供判断忙、完成序号、故障和位置。 *)
END_VAR
VAR_IN_OUT
    awRx : ARRAY[0..31] OF WORD; (* v2 接收字：0=版本2，1=序号，2=命令2启动/3停止；3/4 保留且必须为0，不接受模式写入。 *)
    awTx : ARRAY[0..127] OF WORD; (* 发布字缓冲区 0..127；包含确认、状态、报警、计数和位置，详见程序内索引注释。 *)
END_VAR
VAR_OUTPUT
    xRequest : BOOL; (* 解析到一帧合法新命令时给整机的单扫描请求。 *)
    wRequestSequence : WORD; (* 解析出的新命令序号，供整机处理后原样确认。 *)
    stCommand : ST_RemoteCommand; (* 合法新帧产生的单扫描远程启停请求，没有模式字段。 *)
    uiParseResult : UINT; (* 帧格式检查结果：0 合法，2 版本/模式/命令码不合法，非法帧不下发。 *)
END_VAR
VAR
    aSnapshot : ARRAY[0..31] OF WORD; (* 新命令帧快照，读取后再次核对序号，降低写入过程中读取半帧的风险。 *)
    wLastSeen : WORD; (* 已观察过的帧序号，包含非法帧；相同序号不会重复处理。 *)
    xWasEnabled : BOOL; (* 上扫描通信使能状态；首次使能只记录序号，不执行缓冲区旧命令。 *)
    i : INT; (* 本扫描数组遍历索引；含义及范围以当前 FOR 循环为准。 *)
END_VAR

(* 每扫描清除远程启停脉冲；模式、初始化、复位不属于远程命令。 *)
xRequest:=FALSE;
stCommand.xStart:=FALSE;
stCommand.xStop:=FALSE;
IF NOT xEnable OR NOT xWasEnabled THEN
    (* 首次启用仅记录当前序号，避免重新连接时执行缓冲区遗留命令。 *)
    wLastSeen:=awRx[1];
ELSIF (awRx[1]<>0) AND (awRx[1]<>wLastSeen) THEN
    (* v2：0=版本2，1=新序号，2=命令2启动/3停止，3/4 必须0；旧版或带模式的帧被拒绝。 *)
    aSnapshot:=awRx;
    IF aSnapshot[1]=awRx[1] THEN
        wLastSeen:=aSnapshot[1]; wRequestSequence:=aSnapshot[1]; uiParseResult:=0;
        IF (aSnapshot[0]<>2) OR (aSnapshot[3]<>0) OR (aSnapshot[4]<>0)
           OR ((aSnapshot[2]<>2) AND (aSnapshot[2]<>3)) THEN
            uiParseResult:=2;
        ELSE
            (* 合法新帧只产生启停请求，实际接受还须整机检查本地授权、旋钮模式及状态。 *)
            CASE aSnapshot[2] OF
            2: stCommand.xStart:=TRUE;
            3: stCommand.xStop:=TRUE;
            END_CASE
            xRequest:=TRUE;
        END_IF
    END_IF
END_IF
xWasEnabled:=xEnable;
(* 发布缓冲区是只读反馈，实际寄存器地址与参数下发映射尚未接入。 *)
FOR i:=0 TO 127 DO awTx[i]:=0; END_FOR
(* 0=协议版本2；1=整机处理序号；2=处理结果。 *)
awTx[0]:=2; awTx[1]:=stStatus.wRemoteAckSequence; awTx[2]:=UINT_TO_WORD(stStatus.uiRemoteResult);
(* 3=整机状态；4=自动主步骤。 *)
awTx[3]:=TO_WORD(stStatus.eState); awTx[4]:=TO_WORD(stStatus.eAutoStep);
(* 5/6=报警低字/高字；7/8=循环计数低字/高字。 *)
awTx[5]:=UDINT_TO_WORD(stStatus.udiAlarm); awTx[6]:=UDINT_TO_WORD(SHR(stStatus.udiAlarm,16));
awTx[7]:=UDINT_TO_WORD(stStatus.udiCycleCount); awTx[8]:=UDINT_TO_WORD(SHR(stStatus.udiCycleCount,16));
(* 9=仿真；10=已初始化；11=料到位；12=运行料型。 *)
awTx[9]:=BOOL_TO_WORD(stStatus.xSimulation); awTx[10]:=BOOL_TO_WORD(stStatus.xInitialized);
awTx[11]:=BOOL_TO_WORD(stStatus.xMaterialAtLength); awTx[12]:=UINT_TO_WORD(stStatus.uiActiveMaterialModel);
(* 13=解析器观察序号；14=格式结果0合法/2非法；15=实体旋钮模式0手动/1自动；16=远程启停授权。 *)
awTx[13]:=wRequestSequence; awTx[14]:=UINT_TO_WORD(uiParseResult);
awTx[15]:=TO_WORD(stStatus.eMode);
awTx[16]:=BOOL_TO_WORD(stStatus.xRemoteStartStopAllowed);
(* 17=真实设备接管掩码；18=安全来源0仿真/1真实/2调试旁路；19=是否相对验证；20=初始化拒绝原因。 *)
(* 上位机不能只看 xSimulation：混跑时它恒为 TRUE，必须结合 17 号字判断哪些编号已接实机。 *)
awTx[17]:=stStatus.wRealDeviceMask; awTx[18]:=UINT_TO_WORD(stStatus.uiSafetySource);
awTx[19]:=BOOL_TO_WORD(stStatus.xRelativeVerify); awTx[20]:=UINT_TO_WORD(stStatus.uiInitReject);
(* awTx[32..48]：设备 1..17 位置，按 0.1 工程单位缩放，解读为有符号 INT。 *)
FOR i:=1 TO 17 DO awTx[31+i]:=INT_TO_WORD(LREAL_TO_INT(aStatus[i].lrPosition*10.0)); END_FOR

END_FUNCTION_BLOCK

// Device/Application/04_Machine/FB_IOMap
FUNCTION_BLOCK FB_IOMap
(* 模块说明：设备输出到物理 I/O 的唯一下沉点。真实气缸的阀电平在此写到 GVL_IO_Physical，
   同时仍维护逻辑输出数组供诊断观察。G2 三个侧挡阀在这里按料型逐路下沉。 *)
VAR_INPUT
    aCommand : ARRAY[1..17] OF ST_DeviceCommand; (* 最终设备命令，当前仅用于诊断，不直接驱动输出。 *)
    aStatus : ARRAY[1..17] OF ST_DeviceStatus; (* 各设备的反馈数组 1..17，供判断忙、完成序号、故障和位置。 *)
    aValveOut : ARRAY[1..17] OF BOOL; (* 设备管理器给出的阀电气电平 1..17，真实气缸在此下沉到物理点。 *)
    aValveOutAux : ARRAY[1..17] OF BOOL; (* 第二个执行器的阀电气电平 1..17；G1 右压板在此下沉到物理点。 *)
    aG2Valve : ARRAY[1..3] OF BOOL; (* G2 三个侧挡阀电气电平 1=300，2=450，3=600。 *)
    uiG2Band : UINT; (* G2 当前实际下降的料型带号 300/450/600；0 表示三缸全部提升。 *)
END_VAR
VAR_IN_OUT
    axOutputs : ARRAY[0..31] OF BOOL; (* 逻辑数字输出数组 0..31，按阀电平填写，供在线监视与后续扩展。 *)
END_VAR
VAR
    i : INT; (* 本扫描数组遍历索引；含义及范围以当前 FOR 循环为准。 *)
END_VAR

(* 逻辑输出先清零，只由下面明确赋值的位置置位；未被接管的气缸输出保持失电。 *)
FOR i:=0 TO 31 DO axOutputs[i]:=FALSE; END_FOR

(* ===== 1. 真实气缸阀输出：直接写物理映射符号，TRUE=阀得电=设备动作 ===== *)
(* 未接管时 aValveOut / aG2Valve 为 FALSE，物理点随之失电，不会带着上一个状态一直通电。 *)
GVL_IO_Physical.xDoG1ValveL := aValveOut[9];
GVL_IO_Physical.xDoG1ValveR := aValveOutAux[9];
GVL_IO_Physical.xDoG2Valve300 := aG2Valve[1];
GVL_IO_Physical.xDoG2Valve450 := aG2Valve[2];
GVL_IO_Physical.xDoG2Valve600 := aG2Valve[3];
GVL_IO_Physical.xDoG3Valve := aValveOut[11];
GVL_IO_Physical.xDoG9Valve := aValveOut[17];

(* ===== 2. G2 当前料型带号：供诊断观察，不再从下降反馈反推 ===== *)
GVL_IO.uiG2BandActive := uiG2Band;

(* ===== 3. 逻辑输出镜像：便于在监视表按索引观察，不直接对应物理点 ===== *)
axOutputs[0] := aValveOut[9];
axOutputs[1] := aG2Valve[1];
axOutputs[2] := aG2Valve[2];
axOutputs[3] := aG2Valve[3];
axOutputs[4] := aValveOut[11];
axOutputs[5] := aValveOut[17];

END_FUNCTION_BLOCK

// Device/Application/04_Machine/FB_Indicator
(* 模块说明：面板两色指示灯的纯输出逻辑。指示灯没有反馈、不参与互锁、不占设备索引，
   所以不做成设备，只在这里按整机状态算出两个灯的电平，由 PLC_PRG 下沉到 GVL_IO_Physical。
   优先级：停止/故障最高（红亮绿灭）→ 自动循环运行中（绿慢闪）→ 其余正常运行（绿常亮）。 *)
FUNCTION_BLOCK FB_Indicator
VAR_INPUT
	xRunState : BOOL; (* 整机运行态锁存；FALSE 表示按过停止或上电还没启动。 *)
	eState : E_MachineState; (* 整机状态；Stopped 与 Fault 一律按停机处理。 *)
	eMode : E_MachineMode; (* 模式旋钮当前选择；只有自动循环真正在跑时绿灯才改为慢闪。 *)
	udiAlarm : UDINT; (* 锁存报警码；非 0 时按故障处理，红亮绿灭。 *)
	tBlinkHalf : TIME := T#500MS; (* 慢闪半周期：500 ms 亮 + 500 ms 灭，即每秒亮灭一次。 *)
END_VAR
VAR_OUTPUT
	xGreen : BOOL; (* 绿灯电气电平，TRUE 为亮。 *)
	xRed : BOOL; (* 红灯电气电平，TRUE 为亮。 *)
	xBlinking : BOOL; (* 绿灯当前处于闪烁状态；仅用于监控，不参与控制。 *)
END_VAR
VAR
	tonBlink : TON; (* 闪烁节拍定时器；到点翻转相位并自复位，形成连续方波。 *)
	xBlinkPhase : BOOL; (* 闪烁相位：TRUE 为亮的那一半。 *)
END_VAR

(* 先算闪烁节拍：定时器到点就翻转相位并自复位，得到占空比 50% 的连续方波。
   IN 取 Q 的反相做自复位，Q 每次只保持一个扫描，正好当翻转脉冲用。 *)
tonBlink(IN := NOT tonBlink.Q, PT := tBlinkHalf);
IF tonBlink.Q THEN xBlinkPhase := NOT xBlinkPhase; END_IF

(* 停机判据与状态机保持同一口径：运行态锁存为假、处在故障、或有锁存报警，都算停下。
   红灯优先，任何情况下都不会出现红绿同时亮。 *)
IF (NOT xRunState) OR (eState = E_MachineState.Fault) OR (udiAlarm <> 0) THEN
	xRed := TRUE; xGreen := FALSE; xBlinking := FALSE;
(* 自动循环运行中：绿灯慢闪，表示"正在自动动作"，与手动时有人在场操作区分开。 *)
ELSIF (eMode = E_MachineMode.Automatic) AND (eState = E_MachineState.Automatic) THEN
	xRed := FALSE; xGreen := xBlinkPhase; xBlinking := TRUE;
(* 其余运行状态（手动、初始化中、已就绪待启动）：绿灯常亮。 *)
ELSE
	xRed := FALSE; xGreen := TRUE; xBlinking := FALSE;
END_IF

END_FUNCTION_BLOCK

// Device/Application/90_Legacy/PRG_AxisDemo
(* 模块说明：保留的旧单轴低速往返 Demo，当前未周期调用。它不属于新切割机自动工序。 *)
PROGRAM PRG_AxisDemo
VAR
    (* 运动控制功能块：伺服使能、复位、停止及位置反馈。 *)
    fbPower    : MC_Power; (* 旧 Demo 伺服使能功能块，操作对象为 pandao。 *)
    fbReset    : MC_Reset; (* 旧 Demo 轴故障复位功能块。 *)
    fbStop     : MC_Stop; (* 旧 Demo 受控停止功能块，完成后释放停止锁定。 *)
    fbJog      : MC_Jog; (* 保留的点动实例，当前 Demo 正文未调用。 *)
    fbMoveRel  : MC_MoveRelative; (* 保留的相对定位实例，当前正文使用 fbCycle 执行往返。 *)
    fbMoveAbs  : MC_MoveAbsolute; (* 保留的绝对定位实例，当前 Demo 正文未调用。 *)
    fbCycle    : MC_MoveRelative; (* 实际执行单次往返的相对定位实例，每段使用独立 Execute 触发。 *)
    fbReadPos  : MC_ReadActualPosition; (* 读取 pandao 实际位置，写入旧监控变量 rActPos。 *)
    fbReadStat : MC_ReadStatus; (* 保留的轴状态读取实例，当前正文未调用。 *)
    fbReadErr  : MC_ReadAxisError; (* 保留的轴错误读取实例，当前正文未调用。 *)

    (* 启动信号上升沿检测 *)
    rtCycle    : R_TRIG; (* 旧 Demo 启动按钮上升沿检测，按住按钮不会重复往返。 *)

    (* 自动测试循环的内部状态 *)
    fbCycleExec: BOOL; (* 往返定位功能块 Execute 请求，换向前清除后再置位。 *)
    rCycleDist : LREAL; (* 本段相对位移，正向为正、回程为负，单段绝对值限 20 mm。 *)
    iCycle     : INT := 0; (* 旧 Demo 步骤：0 待机，10 正向，20 停留，30 回程，40 停留结束，99 故障。 *)
    tonDwell   : TON; (* 正向与回程到位后的停留计时器。 *)

    (* 运行状态与故障诊断 *)
    eLastErr   : SMC_ERROR; (* 历史保留的错误变量，当前正文未更新，请看轴/功能块实际错误输出。 *)
	xDoReset: BOOL; (* 历史测试保留变量，当前正文未引用。 *)
	xStopRun: BOOL; (* 旧 Demo 停止请求锁存，收到停止或运动错误后置位。 *)
	rRunDec: LREAL; (* 历史测试保留减速度变量，当前正文未引用。 *)
	xStartRun: BOOL; (* 历史测试保留启动变量，当前正文未引用。 *)
	iStep: INT; (* 历史测试保留步骤变量，当前有效步骤为 iCycle。 *)
	fbMoveVel: MC_MoveVelocity; (* 历史速度运动实例，当前正文未调用。 *)
	Axis: INT; (* 历史保留 INT 变量，不是 pandao 运动轴对象，当前正文未引用。 *)
	Execute: BOOL; (* 历史测试保留执行变量，当前正文未引用。 *)
	rRunVel: LREAL; (* 历史测试保留速度变量，当前正文未引用。 *)
	rRunAcc: LREAL; (* 历史测试保留加速度变量，当前正文未引用。 *)
	Velocity: INT; (* 历史测试保留 INT 变量，当前正文未引用。 *)
	Acceleration: INT; (* 历史测试保留 INT 变量，当前正文未引用。 *)
	Deceleration: INT; (* 历史测试保留 INT 变量，当前正文未引用。 *)
	Direction: INT; (* 历史测试保留方向变量，当前正文未引用。 *)
	InVelocity: INT; (* 历史测试保留 INT 变量，当前正文未引用。 *)
	xMoveExec: BOOL; (* 历史测试保留执行变量，当前正文未引用。 *)
END_VAR

(* 中文注释显示核对：单次低速 20 mm 往返测试。
   GVL_Motion.xStartCycle 的上升沿启动一次循环。
   单程距离最多 20 mm，速度最多 10 mm/s。 *)
rtCycle(CLK := GVL_Motion.xStartCycle);

fbPower(Axis         := pandao,
        Enable       := GVL_Motion.xEnable,
        bRegulatorOn := TRUE,
        bDriveStart  := TRUE);

fbReset(Axis := pandao, Execute := GVL_Motion.xReset);

IF GVL_Motion.xStop THEN
    xStopRun   := TRUE;
    fbCycleExec := FALSE;
    iCycle      := 0;
END_IF

IF fbPower.Error OR fbCycle.Error OR fbReset.Error OR fbStop.Error THEN
    iCycle      := 99;
    fbCycleExec := FALSE;
    xStopRun    := TRUE;
END_IF

fbStop(Axis         := pandao,
       Execute      := xStopRun,
       Deceleration := MIN(MAX(GVL_Motion.rDec, 10.0), 200.0));

IF xStopRun AND fbStop.Done THEN
    xStopRun := FALSE;
END_IF

tonDwell(IN := (iCycle = 20) OR (iCycle = 40),
         PT := GVL_Motion.tDwell);

CASE iCycle OF
    0:  (* 等待启动：一次上升沿触发一次完整往返。 *)
        fbCycleExec := FALSE;
        IF rtCycle.Q
           AND GVL_Motion.xEnable
           AND fbPower.Status
           AND NOT GVL_Motion.xAxisError
           AND NOT xStopRun
           AND (ABS(GVL_Motion.rStroke) > 0.0) THEN
            rCycleDist := MIN(ABS(GVL_Motion.rStroke), 20.0);
            fbCycleExec := TRUE;
            iCycle := 10;
        END_IF

    10: (* 正向运动：等待轴到达指定位置。 *)
        IF fbCycle.Done THEN
            fbCycleExec := FALSE;
            iCycle := 20;
        ELSIF fbCycle.Error THEN
            fbCycleExec := FALSE;
            iCycle := 99;
            xStopRun := TRUE;
        END_IF

    20: (* 正向到位后停留，再发出反向运动指令。 *)
        IF tonDwell.Q AND NOT xStopRun THEN
            rCycleDist := -MIN(ABS(GVL_Motion.rStroke), 20.0);
            fbCycleExec := TRUE;
            iCycle := 30;
        END_IF

    30: (* 反向返回：等待轴完成回程。 *)
        IF fbCycle.Done THEN
            fbCycleExec := FALSE;
            iCycle := 40;
        ELSIF fbCycle.Error THEN
            fbCycleExec := FALSE;
            iCycle := 99;
            xStopRun := TRUE;
        END_IF

    40: (* 返回起点后停留，本次循环结束。 *)
        IF tonDwell.Q THEN
            iCycle := 0;
        END_IF

    99: (* 故障保持：复位成功且停止完成后，允许回到待机。 *)
        fbCycleExec := FALSE;
        IF GVL_Motion.xReset AND fbReset.Done AND NOT xStopRun THEN
            iCycle := 0;
        END_IF

ELSE
    iCycle := 99;
    fbCycleExec := FALSE;
    xStopRun := TRUE;
END_CASE

fbCycle(Axis         := pandao,
        Execute      := fbCycleExec AND NOT xStopRun,
        Distance     := rCycleDist,
        Velocity     := MIN(MAX(GVL_Motion.rVel, 1.0), 10.0),
        Acceleration := MIN(MAX(GVL_Motion.rAcc, 10.0), 200.0),
        Deceleration := MIN(MAX(GVL_Motion.rDec, 10.0), 200.0));

fbReadPos(Axis := pandao, Enable := TRUE);

GVL_Motion.xPowered    := fbPower.Status;
GVL_Motion.xBusy       := fbCycle.Busy OR fbStop.Busy;
GVL_Motion.xDisabled   := NOT fbPower.Status;
GVL_Motion.xStopping   := fbStop.Busy;
GVL_Motion.xStandStill := fbPower.Status AND NOT GVL_Motion.xBusy;
GVL_Motion.xAxisReady  := GVL_Motion.xStandStill AND NOT GVL_Motion.xAxisError;
GVL_Motion.xAxisError  := fbPower.Error OR fbCycle.Error OR fbReset.Error OR fbStop.Error;
GVL_Motion.xErrorStop  := GVL_Motion.xAxisError;
GVL_Motion.iState      := iCycle;
GVL_Motion.rActPos     := fbReadPos.Position;

END_PROGRAM
